TYPE DFC_rbr_outK62SCG : STRUCT
  DTC : UDINT := 16#043C00;
  DFCid : UINT := 682;
  debounceMethod : USINT := TIME_UP_DOWN;
END_STRUCT;
END_TYPE

TYPE DFC_rbr_outK62OR : STRUCT
  DTC : UDINT := 16#043A00;
  DFCid : UINT := 680;
  debounceMethod : USINT := TIME_UP_DOWN;
END_STRUCT;
END_TYPE

TYPE DFC_rbr_safoutChnl1 : STRUCT
  DTC : UDINT := 16#200800;
  DFCid : UINT := 1073;
  debounceMethod : USINT := NO_DEBOUNCE;
END_STRUCT;
END_TYPE

TYPE DFC_rbr_safoutChnl2 : STRUCT
  DTC : UDINT := 16#200900;
  DFCid : UINT := 1103;
  debounceMethod : USINT := NO_DEBOUNCE;
END_STRUCT;
END_TYPE

TYPE DFC_rbr_safoutChnl3 : STRUCT
  DTC : UDINT := 16#200A00;
  DFCid : UINT := 1106;
  debounceMethod : USINT := NO_DEBOUNCE;
END_STRUCT;
END_TYPE

TYPE DFC_rbr_safoutChnl4 : STRUCT
  DTC : UDINT := 16#200B00;
  DFCid : UINT := 1109;
  debounceMethod : USINT := NO_DEBOUNCE;
END_STRUCT;
END_TYPE

TYPE DFC_rbr_safoutChnl5 : STRUCT
  DTC : UDINT := 16#200C00;
  DFCid : UINT := 1112;
  debounceMethod : USINT := NO_DEBOUNCE;
END_STRUCT;
END_TYPE

TYPE DFC_rbr_safoutChnl6 : STRUCT
  DTC : UDINT := 16#201900;
  DFCid : UINT := 1115;
  debounceMethod : USINT := NO_DEBOUNCE;
END_STRUCT;
END_TYPE

TYPE DFC_rbr_safoutChnl7 : STRUCT
  DTC : UDINT := 16#201A00;
  DFCid : UINT := 1118;
  debounceMethod : USINT := NO_DEBOUNCE;
END_STRUCT;
END_TYPE

TYPE DFC_rbr_safoutChnl8 : STRUCT
  DTC : UDINT := 16#201B00;
  DFCid : UINT := 1121;
  debounceMethod : USINT := NO_DEBOUNCE;
END_STRUCT;
END_TYPE

TYPE DFC_rbr_safoutChnl9 : STRUCT
  DTC : UDINT := 16#201C00;
  DFCid : UINT := 1124;
  debounceMethod : USINT := NO_DEBOUNCE;
END_STRUCT;
END_TYPE

TYPE DFC_rbr_safoutChnl10 : STRUCT
  DTC : UDINT := 16#201D00;
  DFCid : UINT := 1074;
  debounceMethod : USINT := NO_DEBOUNCE;
END_STRUCT;
END_TYPE

TYPE DFC_rbr_safoutChnl11 : STRUCT
  DTC : UDINT := 16#201E00;
  DFCid : UINT := 1077;
  debounceMethod : USINT := NO_DEBOUNCE;
END_STRUCT;
END_TYPE

TYPE DFC_rbr_safoutChnl12 : STRUCT
  DTC : UDINT := 16#201F00;
  DFCid : UINT := 1080;
  debounceMethod : USINT := NO_DEBOUNCE;
END_STRUCT;
END_TYPE

TYPE DFC_rbr_safoutChnl13 : STRUCT
  DTC : UDINT := 16#202000;
  DFCid : UINT := 1083;
  debounceMethod : USINT := NO_DEBOUNCE;
END_STRUCT;
END_TYPE

TYPE DFC_rbr_safoutChnl14 : STRUCT
  DTC : UDINT := 16#202100;
  DFCid : UINT := 1086;
  debounceMethod : USINT := NO_DEBOUNCE;
END_STRUCT;
END_TYPE

TYPE DFC_rbr_safoutChnl15 : STRUCT
  DTC : UDINT := 16#202200;
  DFCid : UINT := 1089;
  debounceMethod : USINT := NO_DEBOUNCE;
END_STRUCT;
END_TYPE

TYPE DFC_rbr_safoutChnl16 : STRUCT
  DTC : UDINT := 16#202300;
  DFCid : UINT := 1092;
  debounceMethod : USINT := NO_DEBOUNCE;
END_STRUCT;
END_TYPE

TYPE DFC_rbr_safoutChnl17 : STRUCT
  DTC : UDINT := 16#202400;
  DFCid : UINT := 1095;
  debounceMethod : USINT := NO_DEBOUNCE;
END_STRUCT;
END_TYPE

TYPE DFC_rbr_safoutChnl18 : STRUCT
  DTC : UDINT := 16#202500;
  DFCid : UINT := 1098;
  debounceMethod : USINT := NO_DEBOUNCE;
END_STRUCT;
END_TYPE

TYPE DFC_rbr_safoutChnl6Dev : STRUCT
  DTC : UDINT := 16#202600;
  DFCid : UINT := 1116;
  debounceMethod : USINT := NO_DEBOUNCE;
END_STRUCT;
END_TYPE

TYPE DFC_rbr_safoutChnl7Dev : STRUCT
  DTC : UDINT := 16#202700;
  DFCid : UINT := 1119;
  debounceMethod : USINT := NO_DEBOUNCE;
END_STRUCT;
END_TYPE

TYPE DFC_rbr_safoutChnl8Dev : STRUCT
  DTC : UDINT := 16#202800;
  DFCid : UINT := 1122;
  debounceMethod : USINT := NO_DEBOUNCE;
END_STRUCT;
END_TYPE

TYPE DFC_rbr_safoutChnl9Dev : STRUCT
  DTC : UDINT := 16#202900;
  DFCid : UINT := 1125;
  debounceMethod : USINT := NO_DEBOUNCE;
END_STRUCT;
END_TYPE

TYPE DFC_rbr_safoutChnl10Dev : STRUCT
  DTC : UDINT := 16#202A00;
  DFCid : UINT := 1075;
  debounceMethod : USINT := NO_DEBOUNCE;
END_STRUCT;
END_TYPE

TYPE DFC_rbr_safoutChnl11Dev : STRUCT
  DTC : UDINT := 16#202B00;
  DFCid : UINT := 1078;
  debounceMethod : USINT := NO_DEBOUNCE;
END_STRUCT;
END_TYPE

TYPE DFC_rbr_safoutChnl12Dev : STRUCT
  DTC : UDINT := 16#202C00;
  DFCid : UINT := 1081;
  debounceMethod : USINT := NO_DEBOUNCE;
END_STRUCT;
END_TYPE

TYPE DFC_rbr_safoutChnl13Dev : STRUCT
  DTC : UDINT := 16#202D00;
  DFCid : UINT := 1084;
  debounceMethod : USINT := NO_DEBOUNCE;
END_STRUCT;
END_TYPE

TYPE DFC_rbr_safoutChnl14Dev : STRUCT
  DTC : UDINT := 16#202E00;
  DFCid : UINT := 1087;
  debounceMethod : USINT := NO_DEBOUNCE;
END_STRUCT;
END_TYPE

TYPE DFC_rbr_safoutChnl15Dev : STRUCT
  DTC : UDINT := 16#202F00;
  DFCid : UINT := 1090;
  debounceMethod : USINT := NO_DEBOUNCE;
END_STRUCT;
END_TYPE

TYPE DFC_rbr_safoutChnl16Dev : STRUCT
  DTC : UDINT := 16#203000;
  DFCid : UINT := 1093;
  debounceMethod : USINT := NO_DEBOUNCE;
END_STRUCT;
END_TYPE

TYPE DFC_rbr_safoutChnl17Dev : STRUCT
  DTC : UDINT := 16#203100;
  DFCid : UINT := 1096;
  debounceMethod : USINT := NO_DEBOUNCE;
END_STRUCT;
END_TYPE

TYPE DFC_rbr_safoutChnl18Dev : STRUCT
  DTC : UDINT := 16#203200;
  DFCid : UINT := 1099;
  debounceMethod : USINT := NO_DEBOUNCE;
END_STRUCT;
END_TYPE

TYPE DFC_rbr_safoutChnl1OR : STRUCT
  DTC : UDINT := 16#200D00;
  DFCid : UINT := 1102;
  debounceMethod : USINT := NO_DEBOUNCE;
END_STRUCT;
END_TYPE

TYPE DFC_rbr_safoutChnl2OR : STRUCT
  DTC : UDINT := 16#200E00;
  DFCid : UINT := 1105;
  debounceMethod : USINT := NO_DEBOUNCE;
END_STRUCT;
END_TYPE

TYPE DFC_rbr_safoutChnl3OR : STRUCT
  DTC : UDINT := 16#200F00;
  DFCid : UINT := 1108;
  debounceMethod : USINT := NO_DEBOUNCE;
END_STRUCT;
END_TYPE

TYPE DFC_rbr_safoutChnl4OR : STRUCT
  DTC : UDINT := 16#201100;
  DFCid : UINT := 1111;
  debounceMethod : USINT := NO_DEBOUNCE;
END_STRUCT;
END_TYPE

TYPE DFC_rbr_safoutChnl5OR : STRUCT
  DTC : UDINT := 16#201200;
  DFCid : UINT := 1114;
  debounceMethod : USINT := NO_DEBOUNCE;
END_STRUCT;
END_TYPE

TYPE DFC_rbr_safoutChnl6OR : STRUCT
  DTC : UDINT := 16#203300;
  DFCid : UINT := 1117;
  debounceMethod : USINT := NO_DEBOUNCE;
END_STRUCT;
END_TYPE

TYPE DFC_rbr_safoutChnl7OR : STRUCT
  DTC : UDINT := 16#203400;
  DFCid : UINT := 1120;
  debounceMethod : USINT := NO_DEBOUNCE;
END_STRUCT;
END_TYPE

TYPE DFC_rbr_safoutChnl8OR : STRUCT
  DTC : UDINT := 16#203500;
  DFCid : UINT := 1123;
  debounceMethod : USINT := NO_DEBOUNCE;
END_STRUCT;
END_TYPE

TYPE DFC_rbr_safoutChnl9OR : STRUCT
  DTC : UDINT := 16#203600;
  DFCid : UINT := 1126;
  debounceMethod : USINT := NO_DEBOUNCE;
END_STRUCT;
END_TYPE

TYPE DFC_rbr_safoutChnl10OR : STRUCT
  DTC : UDINT := 16#203700;
  DFCid : UINT := 1076;
  debounceMethod : USINT := NO_DEBOUNCE;
END_STRUCT;
END_TYPE

TYPE DFC_rbr_safoutChnl11OR : STRUCT
  DTC : UDINT := 16#203800;
  DFCid : UINT := 1079;
  debounceMethod : USINT := NO_DEBOUNCE;
END_STRUCT;
END_TYPE

TYPE DFC_rbr_safoutChnl12OR : STRUCT
  DTC : UDINT := 16#203900;
  DFCid : UINT := 1082;
  debounceMethod : USINT := NO_DEBOUNCE;
END_STRUCT;
END_TYPE

TYPE DFC_rbr_safoutChnl13OR : STRUCT
  DTC : UDINT := 16#203A00;
  DFCid : UINT := 1085;
  debounceMethod : USINT := NO_DEBOUNCE;
END_STRUCT;
END_TYPE

TYPE DFC_rbr_safoutChnl14OR : STRUCT
  DTC : UDINT := 16#203B00;
  DFCid : UINT := 1088;
  debounceMethod : USINT := NO_DEBOUNCE;
END_STRUCT;
END_TYPE

TYPE DFC_rbr_safoutChnl15OR : STRUCT
  DTC : UDINT := 16#203C00;
  DFCid : UINT := 1091;
  debounceMethod : USINT := NO_DEBOUNCE;
END_STRUCT;
END_TYPE

TYPE DFC_rbr_safoutChnl16OR : STRUCT
  DTC : UDINT := 16#203D00;
  DFCid : UINT := 1094;
  debounceMethod : USINT := NO_DEBOUNCE;
END_STRUCT;
END_TYPE

TYPE DFC_rbr_safoutChnl17OR : STRUCT
  DTC : UDINT := 16#203E00;
  DFCid : UINT := 1097;
  debounceMethod : USINT := NO_DEBOUNCE;
END_STRUCT;
END_TYPE

TYPE DFC_rbr_safoutChnl18OR : STRUCT
  DTC : UDINT := 16#203F00;
  DFCid : UINT := 1100;
  debounceMethod : USINT := NO_DEBOUNCE;
END_STRUCT;
END_TYPE

TYPE DFC_rbr_safoutCfg : STRUCT
  DTC : UDINT := 16#200100;
  DFCid : UINT := 1072;
  debounceMethod : USINT := NO_DEBOUNCE;
END_STRUCT;
END_TYPE

TYPE DFC_rbr_safout : STRUCT
  DTC : UDINT := 16#200200;
  DFCid : UINT := 1071;
  debounceMethod : USINT := NO_DEBOUNCE;
END_STRUCT;
END_TYPE

TYPE DFC_rbr_safoutGetStatus : STRUCT
  DTC : UDINT := 16#200300;
  DFCid : UINT := 1128;
  debounceMethod : USINT := NO_DEBOUNCE;
END_STRUCT;
END_TYPE

TYPE DFC_rbr_safoutDevError : STRUCT
  DTC : UDINT := 16#201800;
  DFCid : UINT := 1127;
  debounceMethod : USINT := NO_DEBOUNCE;
END_STRUCT;
END_TYPE

TYPE DFC_rbr_safoutResetError : STRUCT
  DTC : UDINT := 16#200400;
  DFCid : UINT := 1130;
  debounceMethod : USINT := NO_DEBOUNCE;
END_STRUCT;
END_TYPE

TYPE DFC_rbr_safoutIgnoreError : STRUCT
  DTC : UDINT := 16#200500;
  DFCid : UINT := 1129;
  debounceMethod : USINT := NO_DEBOUNCE;
END_STRUCT;
END_TYPE

TYPE DFC_rbr_safoutUnlock : STRUCT
  DTC : UDINT := 16#200600;
  DFCid : UINT := 1131;
  debounceMethod : USINT := NO_DEBOUNCE;
END_STRUCT;
END_TYPE

TYPE DFC_rbr_outDo : STRUCT
  DTC : UDINT := 16#048300;
  DFCid : UINT := 1025;
  debounceMethod : USINT := NO_DEBOUNCE;
END_STRUCT;
END_TYPE

TYPE DFC_rbr_outDoGetCurrent : STRUCT
  DTC : UDINT := 16#048400;
  DFCid : UINT := 1028;
  debounceMethod : USINT := NO_DEBOUNCE;
END_STRUCT;
END_TYPE

TYPE DFC_rbr_outPod : STRUCT
  DTC : UDINT := 16#048B00;
  DFCid : UINT := 1067;
  debounceMethod : USINT := NO_DEBOUNCE;
END_STRUCT;
END_TYPE

TYPE DFC_rbr_outPodCfg : STRUCT
  DTC : UDINT := 16#048C00;
  DFCid : UINT := 1068;
  debounceMethod : USINT := NO_DEBOUNCE;
END_STRUCT;
END_TYPE

TYPE DFC_rbr_outPodCfgPeriod : STRUCT
  DTC : UDINT := 16#048D00;
  DFCid : UINT := 1069;
  debounceMethod : USINT := NO_DEBOUNCE;
END_STRUCT;
END_TYPE

TYPE DFC_rbr_outPoc : STRUCT
  DTC : UDINT := 16#048600;
  DFCid : UINT := 1063;
  debounceMethod : USINT := NO_DEBOUNCE;
END_STRUCT;
END_TYPE

TYPE DFC_rbr_outPocCfg : STRUCT
  DTC : UDINT := 16#048800;
  DFCid : UINT := 1064;
  debounceMethod : USINT := NO_DEBOUNCE;
END_STRUCT;
END_TYPE

TYPE DFC_rbr_outPoCfg : STRUCT
  DTC : UDINT := 16#048700;
  DFCid : UINT := 1056;
  debounceMethod : USINT := NO_DEBOUNCE;
END_STRUCT;
END_TYPE

TYPE DFC_rbr_outPocCfgPI : STRUCT
  DTC : UDINT := 16#048A00;
  DFCid : UINT := 1066;
  debounceMethod : USINT := NO_DEBOUNCE;
END_STRUCT;
END_TYPE

TYPE DFC_rbr_outPocCfgDither : STRUCT
  DTC : UDINT := 16#048900;
  DFCid : UINT := 1065;
  debounceMethod : USINT := NO_DEBOUNCE;
END_STRUCT;
END_TYPE

TYPE DFC_rbr_outPoGetCurrent : STRUCT
  DTC : UDINT := 16#048E00;
  DFCid : UINT := 1060;
  debounceMethod : USINT := NO_DEBOUNCE;
END_STRUCT;
END_TYPE

TYPE DFC_rbr_outAov : STRUCT
  DTC : UDINT := 16#048000;
  DFCid : UINT := 1019;
  debounceMethod : USINT := NO_DEBOUNCE;
END_STRUCT;
END_TYPE

TYPE DFC_rbr_outAovCfg : STRUCT
  DTC : UDINT := 16#048100;
  DFCid : UINT := 1020;
  debounceMethod : USINT := NO_DEBOUNCE;
END_STRUCT;
END_TYPE

TYPE DFC_rbr_outAovCfgPI : STRUCT
  DTC : UDINT := 16#14D700;
  DFCid : UINT := 1021;
  debounceMethod : USINT := NO_DEBOUNCE;
END_STRUCT;
END_TYPE

TYPE DFC_rbr_outAovGetVoltage : STRUCT
  DTC : UDINT := 16#048200;
  DFCid : UINT := 1023;
  debounceMethod : USINT := NO_DEBOUNCE;
END_STRUCT;
END_TYPE

TYPE DFC_rbr_outDoGetStatus : STRUCT
  DTC : UDINT := 16#048F00;
  DFCid : UINT := 1029;
  debounceMethod : USINT := NO_DEBOUNCE;
END_STRUCT;
END_TYPE

TYPE DFC_rbr_outDoResetError : STRUCT
  DTC : UDINT := 16#049000;
  DFCid : UINT := 1030;
  debounceMethod : USINT := NO_DEBOUNCE;
END_STRUCT;
END_TYPE

TYPE DFC_rbr_outPo : STRUCT
  DTC : UDINT := 16#049100;
  DFCid : UINT := 1055;
  debounceMethod : USINT := NO_DEBOUNCE;
END_STRUCT;
END_TYPE

TYPE DFC_rbr_outPoCfgPeriod : STRUCT
  DTC : UDINT := 16#049200;
  DFCid : UINT := 1057;
  debounceMethod : USINT := NO_DEBOUNCE;
END_STRUCT;
END_TYPE

TYPE DFC_rbr_outPoGetStatus : STRUCT
  DTC : UDINT := 16#049300;
  DFCid : UINT := 1061;
  debounceMethod : USINT := NO_DEBOUNCE;
END_STRUCT;
END_TYPE

TYPE DFC_rbr_outPoResetError : STRUCT
  DTC : UDINT := 16#049400;
  DFCid : UINT := 1062;
  debounceMethod : USINT := NO_DEBOUNCE;
END_STRUCT;
END_TYPE

TYPE DFC_rbr_outAovGetStatus : STRUCT
  DTC : UDINT := 16#049500;
  DFCid : UINT := 1022;
  debounceMethod : USINT := NO_DEBOUNCE;
END_STRUCT;
END_TYPE

TYPE DFC_rbr_outAovResetError : STRUCT
  DTC : UDINT := 16#049600;
  DFCid : UINT := 1024;
  debounceMethod : USINT := NO_DEBOUNCE;
END_STRUCT;
END_TYPE

TYPE DFC_rbr_sysAiv : STRUCT
  DTC : UDINT := 16#010100;
  DFCid : UINT := 1146;
  debounceMethod : USINT := NO_DEBOUNCE;
END_STRUCT;
END_TYPE

TYPE DFC_rbr_memFlsCfgShr : STRUCT
  DTC : UDINT := 16#060900;
  DFCid : UINT := 953;
  debounceMethod : USINT := NO_DEBOUNCE;
END_STRUCT;
END_TYPE

TYPE DFC_rbr_sysDo : STRUCT
  DTC : UDINT := 16#010200;
  DFCid : UINT := 1148;
  debounceMethod : USINT := NO_DEBOUNCE;
END_STRUCT;
END_TYPE

TYPE DFC_rbr_sysGetVss : STRUCT
  DTC : UDINT := 16#010600;
  DFCid : UINT := 1149;
  debounceMethod : USINT := NO_DEBOUNCE;
END_STRUCT;
END_TYPE

TYPE DFC_rbr_sysDi : STRUCT
  DTC : UDINT := 16#010300;
  DFCid : UINT := 1147;
  debounceMethod : USINT := NO_DEBOUNCE;
END_STRUCT;
END_TYPE

TYPE DFC_rbr_sysAit : STRUCT
  DTC : UDINT := 16#010400;
  DFCid : UINT := 1145;
  debounceMethod : USINT := NO_DEBOUNCE;
END_STRUCT;
END_TYPE

TYPE DFC_rbr_sysSetVss : STRUCT
  DTC : UDINT := 16#010500;
  DFCid : UINT := 1153;
  debounceMethod : USINT := NO_DEBOUNCE;
END_STRUCT;
END_TYPE

TYPE DFC_rbr_outPoDisable : STRUCT
  DTC : UDINT := 16#049800;
  DFCid : UINT := 1059;
  debounceMethod : USINT := NO_DEBOUNCE;
END_STRUCT;
END_TYPE

TYPE DFC_rbr_safout_cfgDiag : STRUCT
  DTC : UDINT := 16#200700;
  DFCid : UINT := 1132;
  debounceMethod : USINT := NO_DEBOUNCE;
END_STRUCT;
END_TYPE

TYPE DFC_rbr_outDoDisable : STRUCT
  DTC : UDINT := 16#049700;
  DFCid : UINT := 1027;
  debounceMethod : USINT := NO_DEBOUNCE;
END_STRUCT;
END_TYPE

TYPE DFC_rbr_sysOperHrIntegrityErr : STRUCT
  DTC : UDINT := 16#010A00;
  DFCid : UINT := 1151;
  debounceMethod : USINT := NO_DEBOUNCE;
END_STRUCT;
END_TYPE

TYPE DFC_rbr_sysOperHrsSaturated : STRUCT
  DTC : UDINT := 16#010B00;
  DFCid : UINT := 1152;
  debounceMethod : USINT := NO_DEBOUNCE;
END_STRUCT;
END_TYPE

TYPE DFC_rbr_mo_INHLatch : STRUCT
  DTC : UDINT := 16#082200;
  DFCid : UINT := 968;
  debounceMethod : USINT := NO_DEBOUNCE;
END_STRUCT;
END_TYPE

TYPE DFC_rbr_mo_INH : STRUCT
  DTC : UDINT := 16#082100;
  DFCid : UINT := 967;
  debounceMethod : USINT := NO_DEBOUNCE;
END_STRUCT;
END_TYPE

TYPE DFC_rbr_memReadSystemError : STRUCT
  DTC : UDINT := 16#060800;
  DFCid : UINT := 961;
  debounceMethod : USINT := NO_DEBOUNCE;
END_STRUCT;
END_TYPE

TYPE DFC_rbr_memReadCalibInputError : STRUCT
  DTC : UDINT := 16#060A00;
  DFCid : UINT := 959;
  debounceMethod : USINT := NO_DEBOUNCE;
END_STRUCT;
END_TYPE

TYPE DFC_rbr_memReadCalibOuputError : STRUCT
  DTC : UDINT := 16#060B00;
  DFCid : UINT := 960;
  debounceMethod : USINT := NO_DEBOUNCE;
END_STRUCT;
END_TYPE

TYPE DFC_rbr_memReadApi2Error : STRUCT
  DTC : UDINT := 16#060600;
  DFCid : UINT := 957;
  debounceMethod : USINT := NO_DEBOUNCE;
END_STRUCT;
END_TYPE

TYPE DFC_rbr_memReadApi1Error : STRUCT
  DTC : UDINT := 16#060500;
  DFCid : UINT := 956;
  debounceMethod : USINT := NO_DEBOUNCE;
END_STRUCT;
END_TYPE

TYPE DFC_rbr_memMarkBlock : STRUCT
  DTC : UDINT := 16#060400;
  DFCid : UINT := 955;
  debounceMethod : USINT := NO_DEBOUNCE;
END_STRUCT;
END_TYPE

TYPE DFC_rbr_safoutChnl3Dev : STRUCT
  DTC : UDINT := 16#201500;
  DFCid : UINT := 1107;
  debounceMethod : USINT := NO_DEBOUNCE;
END_STRUCT;
END_TYPE

TYPE DFC_rbr_safoutChnl5Dev : STRUCT
  DTC : UDINT := 16#201700;
  DFCid : UINT := 1113;
  debounceMethod : USINT := NO_DEBOUNCE;
END_STRUCT;
END_TYPE

TYPE DFC_rbr_safoutChnl4Dev : STRUCT
  DTC : UDINT := 16#201600;
  DFCid : UINT := 1110;
  debounceMethod : USINT := NO_DEBOUNCE;
END_STRUCT;
END_TYPE

TYPE DFC_rbr_safoutChnl2Dev : STRUCT
  DTC : UDINT := 16#201400;
  DFCid : UINT := 1104;
  debounceMethod : USINT := NO_DEBOUNCE;
END_STRUCT;
END_TYPE

TYPE DFC_rbr_safoutChnl1Dev : STRUCT
  DTC : UDINT := 16#201300;
  DFCid : UINT := 1101;
  debounceMethod : USINT := NO_DEBOUNCE;
END_STRUCT;
END_TYPE

TYPE DFC_rbr_outPoCfgPwrLs : STRUCT
  DTC : UDINT := 16#049900;
  DFCid : UINT := 1058;
  debounceMethod : USINT := NO_DEBOUNCE;
END_STRUCT;
END_TYPE

TYPE DFC_rbr_lin_wakeUp : STRUCT
  DTC : UDINT := 16#210000;
  DFCid : UINT := 952;
  debounceMethod : USINT := NO_DEBOUNCE;
END_STRUCT;
END_TYPE

TYPE DFC_rbr_lin_gotoSleep : STRUCT
  DTC : UDINT := 16#210200;
  DFCid : UINT := 950;
  debounceMethod : USINT := NO_DEBOUNCE;
END_STRUCT;
END_TYPE

TYPE DFC_rbr_lin_getStatus : STRUCT
  DTC : UDINT := 16#210300;
  DFCid : UINT := 949;
  debounceMethod : USINT := NO_DEBOUNCE;
END_STRUCT;
END_TYPE

TYPE DFC_rbr_lin_scheduleRequest : STRUCT
  DTC : UDINT := 16#210100;
  DFCid : UINT := 951;
  debounceMethod : USINT := NO_DEBOUNCE;
END_STRUCT;
END_TYPE

TYPE DFC_rbr_lin_SendSignal : STRUCT
  DTC : UDINT := 16#210400;
  DFCid : UINT := 948;
  debounceMethod : USINT := NO_DEBOUNCE;
END_STRUCT;
END_TYPE

TYPE DFC_rbr_inPhaseGetStatus : STRUCT
  DTC : UDINT := 16#039F00;
  DFCid : UINT := 897;
  debounceMethod : USINT := NO_DEBOUNCE;
END_STRUCT;
END_TYPE

TYPE DFC_rbr_inPhaseResetCounter : STRUCT
  DTC : UDINT := 16#03A000;
  DFCid : UINT := 898;
  debounceMethod : USINT := NO_DEBOUNCE;
END_STRUCT;
END_TYPE

TYPE DFC_rbr_inPhase : STRUCT
  DTC : UDINT := 16#039E00;
  DFCid : UINT := 896;
  debounceMethod : USINT := NO_DEBOUNCE;
END_STRUCT;
END_TYPE

TYPE DFC_rbr_inFi_Buffered : STRUCT
  DTC : UDINT := 16#135200;
  DFCid : UINT := 895;
  debounceMethod : USINT := NO_DEBOUNCE;
END_STRUCT;
END_TYPE

TYPE DFC_rbr_secGetLevel : STRUCT
  DTC : UDINT := 16#220200;
  DFCid : UINT := 1137;
  debounceMethod : USINT := NO_DEBOUNCE;
END_STRUCT;
END_TYPE

TYPE DFC_rbr_secSetLevel : STRUCT
  DTC : UDINT := 16#220300;
  DFCid : UINT := 1144;
  debounceMethod : USINT := NO_DEBOUNCE;
END_STRUCT;
END_TYPE

TYPE DFC_rbr_secSaveSecret : STRUCT
  DTC : UDINT := 16#220100;
  DFCid : UINT := 1143;
  debounceMethod : USINT := NO_DEBOUNCE;
END_STRUCT;
END_TYPE

TYPE DFC_rbr_secGetSeed : STRUCT
  DTC : UDINT := 16#220000;
  DFCid : UINT := 1139;
  debounceMethod : USINT := NO_DEBOUNCE;
END_STRUCT;
END_TYPE

TYPE DFC_rbr_secIsRequestAllowed : STRUCT
  DTC : UDINT := 16#220700;
  DFCid : UINT := 1141;
  debounceMethod : USINT := NO_DEBOUNCE;
END_STRUCT;
END_TYPE

TYPE DFC_rbr_secGetRnd : STRUCT
  DTC : UDINT := 16#220600;
  DFCid : UINT := 1138;
  debounceMethod : USINT := NO_DEBOUNCE;
END_STRUCT;
END_TYPE

TYPE DFC_rbr_secEvalRespKey : STRUCT
  DTC : UDINT := 16#220500;
  DFCid : UINT := 1135;
  debounceMethod : USINT := NO_DEBOUNCE;
END_STRUCT;
END_TYPE

TYPE DFC_rbr_secResetLevel : STRUCT
  DTC : UDINT := 16#220400;
  DFCid : UINT := 1142;
  debounceMethod : USINT := NO_DEBOUNCE;
END_STRUCT;
END_TYPE

TYPE DFC_rbr_lin_ReceiveSignal : STRUCT
  DTC : UDINT := 16#210500;
  DFCid : UINT := 947;
  debounceMethod : USINT := NO_DEBOUNCE;
END_STRUCT;
END_TYPE

TYPE DFC_rbr_sys_coreload : STRUCT
  DTC : UDINT := 16#010900;
  DFCid : UINT := 1154;
  debounceMethod : USINT := NO_DEBOUNCE;
END_STRUCT;
END_TYPE

TYPE DFC_rbr_sys_taskload : STRUCT
  DTC : UDINT := 16#010800;
  DFCid : UINT := 1155;
  debounceMethod : USINT := NO_DEBOUNCE;
END_STRUCT;
END_TYPE

TYPE DFC_rbr_dsmDTCJ1939 : STRUCT
  DTC : UDINT := 16#071000;
  DFCid : UINT := 868;
  debounceMethod : USINT := NO_DEBOUNCE;
END_STRUCT;
END_TYPE

TYPE DFC_rbr_sysInit : STRUCT
  DTC : UDINT := 16#010700;
  DFCid : UINT := 1150;
  debounceMethod : USINT := NO_DEBOUNCE;
END_STRUCT;
END_TYPE

TYPE DFC_rbr_outK07Unintended : STRUCT
  DTC : UDINT := 16#14CB00;
  DFCid : UINT := 1032;
  debounceMethod : USINT := NO_DEBOUNCE;
END_STRUCT;
END_TYPE

TYPE DFC_rbr_outK09Unintended : STRUCT
  DTC : UDINT := 16#14CD00;
  DFCid : UINT := 1036;
  debounceMethod : USINT := NO_DEBOUNCE;
END_STRUCT;
END_TYPE

TYPE DFC_rbr_outK73Unintended : STRUCT
  DTC : UDINT := 16#14D600;
  DFCid : UINT := 1054;
  debounceMethod : USINT := NO_DEBOUNCE;
END_STRUCT;
END_TYPE

TYPE DFC_rbr_outK08Unintended : STRUCT
  DTC : UDINT := 16#14CC00;
  DFCid : UINT := 1034;
  debounceMethod : USINT := NO_DEBOUNCE;
END_STRUCT;
END_TYPE

TYPE DFC_rbr_outK29Unintended : STRUCT
  DTC : UDINT := 16#14D400;
  DFCid : UINT := 1050;
  debounceMethod : USINT := NO_DEBOUNCE;
END_STRUCT;
END_TYPE

TYPE DFC_rbr_outK17Unintended : STRUCT
  DTC : UDINT := 16#14D300;
  DFCid : UINT := 1048;
  debounceMethod : USINT := NO_DEBOUNCE;
END_STRUCT;
END_TYPE

TYPE DFC_rbr_outK16Unintended : STRUCT
  DTC : UDINT := 16#14D200;
  DFCid : UINT := 1046;
  debounceMethod : USINT := NO_DEBOUNCE;
END_STRUCT;
END_TYPE

TYPE DFC_rbr_outK14Unintended : STRUCT
  DTC : UDINT := 16#14D000;
  DFCid : UINT := 1042;
  debounceMethod : USINT := NO_DEBOUNCE;
END_STRUCT;
END_TYPE

TYPE DFC_rbr_outK15Unintended : STRUCT
  DTC : UDINT := 16#14D100;
  DFCid : UINT := 1044;
  debounceMethod : USINT := NO_DEBOUNCE;
END_STRUCT;
END_TYPE

TYPE DFC_rbr_outK51Unintended : STRUCT
  DTC : UDINT := 16#14D500;
  DFCid : UINT := 1052;
  debounceMethod : USINT := NO_DEBOUNCE;
END_STRUCT;
END_TYPE

TYPE DFC_rbr_outK12Unintended : STRUCT
  DTC : UDINT := 16#14CE00;
  DFCid : UINT := 1038;
  debounceMethod : USINT := NO_DEBOUNCE;
END_STRUCT;
END_TYPE

TYPE DFC_rbr_outK13Unintended : STRUCT
  DTC : UDINT := 16#14CF00;
  DFCid : UINT := 1040;
  debounceMethod : USINT := NO_DEBOUNCE;
END_STRUCT;
END_TYPE

TYPE DFC_rbr_outA32Unintended : STRUCT
  DTC : UDINT := 16#14C000;
  DFCid : UINT := 998;
  debounceMethod : USINT := NO_DEBOUNCE;
END_STRUCT;
END_TYPE

TYPE DFC_rbr_outA47Unintended : STRUCT
  DTC : UDINT := 16#14C500;
  DFCid : UINT := 1008;
  debounceMethod : USINT := NO_DEBOUNCE;
END_STRUCT;
END_TYPE

TYPE DFC_rbr_outA31Unintended : STRUCT
  DTC : UDINT := 16#14BF00;
  DFCid : UINT := 996;
  debounceMethod : USINT := NO_DEBOUNCE;
END_STRUCT;
END_TYPE

TYPE DFC_rbr_outA48Unintended : STRUCT
  DTC : UDINT := 16#14C600;
  DFCid : UINT := 1010;
  debounceMethod : USINT := NO_DEBOUNCE;
END_STRUCT;
END_TYPE

TYPE DFC_rbr_outA46Unintended : STRUCT
  DTC : UDINT := 16#14C400;
  DFCid : UINT := 1006;
  debounceMethod : USINT := NO_DEBOUNCE;
END_STRUCT;
END_TYPE

TYPE DFC_rbr_outA33Unintended : STRUCT
  DTC : UDINT := 16#14C100;
  DFCid : UINT := 1000;
  debounceMethod : USINT := NO_DEBOUNCE;
END_STRUCT;
END_TYPE

TYPE DFC_rbr_outA19Unintended : STRUCT
  DTC : UDINT := 16#14BD00;
  DFCid : UINT := 992;
  debounceMethod : USINT := NO_DEBOUNCE;
END_STRUCT;
END_TYPE

TYPE DFC_rbr_outA05Unintended : STRUCT
  DTC : UDINT := 16#14B600;
  DFCid : UINT := 978;
  debounceMethod : USINT := NO_DEBOUNCE;
END_STRUCT;
END_TYPE

TYPE DFC_rbr_outA20Unintended : STRUCT
  DTC : UDINT := 16#14BE00;
  DFCid : UINT := 994;
  debounceMethod : USINT := NO_DEBOUNCE;
END_STRUCT;
END_TYPE

TYPE DFC_rbr_outA03Unintended : STRUCT
  DTC : UDINT := 16#14B400;
  DFCid : UINT := 974;
  debounceMethod : USINT := NO_DEBOUNCE;
END_STRUCT;
END_TYPE

TYPE DFC_rbr_outA18Unintended : STRUCT
  DTC : UDINT := 16#14BC00;
  DFCid : UINT := 990;
  debounceMethod : USINT := NO_DEBOUNCE;
END_STRUCT;
END_TYPE

TYPE DFC_rbr_outA04Unintended : STRUCT
  DTC : UDINT := 16#14B500;
  DFCid : UINT := 976;
  debounceMethod : USINT := NO_DEBOUNCE;
END_STRUCT;
END_TYPE

TYPE DFC_rbr_outA34Unintended : STRUCT
  DTC : UDINT := 16#14C200;
  DFCid : UINT := 1002;
  debounceMethod : USINT := NO_DEBOUNCE;
END_STRUCT;
END_TYPE

TYPE DFC_rbr_outA51Unintended : STRUCT
  DTC : UDINT := 16#14C700;
  DFCid : UINT := 1012;
  debounceMethod : USINT := NO_DEBOUNCE;
END_STRUCT;
END_TYPE

TYPE DFC_rbr_outA35Unintended : STRUCT
  DTC : UDINT := 16#14C300;
  DFCid : UINT := 1004;
  debounceMethod : USINT := NO_DEBOUNCE;
END_STRUCT;
END_TYPE

TYPE DFC_rbr_outA53Unintended : STRUCT
  DTC : UDINT := 16#14C900;
  DFCid : UINT := 1016;
  debounceMethod : USINT := NO_DEBOUNCE;
END_STRUCT;
END_TYPE

TYPE DFC_rbr_outA52Unintended : STRUCT
  DTC : UDINT := 16#14C800;
  DFCid : UINT := 1014;
  debounceMethod : USINT := NO_DEBOUNCE;
END_STRUCT;
END_TYPE

TYPE DFC_rbr_outA54Unintended : STRUCT
  DTC : UDINT := 16#14CA00;
  DFCid : UINT := 1018;
  debounceMethod : USINT := NO_DEBOUNCE;
END_STRUCT;
END_TYPE

TYPE DFC_rbr_outA09Unintended : STRUCT
  DTC : UDINT := 16#14B900;
  DFCid : UINT := 984;
  debounceMethod : USINT := NO_DEBOUNCE;
END_STRUCT;
END_TYPE

TYPE DFC_rbr_outA02Unintended : STRUCT
  DTC : UDINT := 16#14B300;
  DFCid : UINT := 972;
  debounceMethod : USINT := NO_DEBOUNCE;
END_STRUCT;
END_TYPE

TYPE DFC_rbr_outA17Unintended : STRUCT
  DTC : UDINT := 16#14BB00;
  DFCid : UINT := 988;
  debounceMethod : USINT := NO_DEBOUNCE;
END_STRUCT;
END_TYPE

TYPE DFC_rbr_outA08Unintended : STRUCT
  DTC : UDINT := 16#14B800;
  DFCid : UINT := 982;
  debounceMethod : USINT := NO_DEBOUNCE;
END_STRUCT;
END_TYPE

TYPE DFC_rbr_outA07Unintended : STRUCT
  DTC : UDINT := 16#14B700;
  DFCid : UINT := 980;
  debounceMethod : USINT := NO_DEBOUNCE;
END_STRUCT;
END_TYPE

TYPE DFC_rbr_outA10Unintended : STRUCT
  DTC : UDINT := 16#14BA00;
  DFCid : UINT := 986;
  debounceMethod : USINT := NO_DEBOUNCE;
END_STRUCT;
END_TYPE

TYPE DFC_rbr_outDoCfgPwrLs : STRUCT
  DTC : UDINT := 16#14D800;
  DFCid : UINT := 1026;
  debounceMethod : USINT := NO_DEBOUNCE;
END_STRUCT;
END_TYPE

TYPE DFC_rbr_mo_memoryProtection_err : STRUCT
  DTC : UDINT := 16#083300;
  DFCid : UINT := 970;
  debounceMethod : USINT := NO_DEBOUNCE;
END_STRUCT;
END_TYPE

TYPE DFC_rbr_rsmFfiApiCallErr : STRUCT
  DTC : UDINT := 16#010C00;
  DFCid : UINT := 1070;
  debounceMethod : USINT := NO_DEBOUNCE;
END_STRUCT;
END_TYPE

TYPE DFC_rbr_isobusSftyCanTxErr : STRUCT
  DTC : UDINT := 16#051F00;
  DFCid : UINT := 946;
  debounceMethod : USINT := NO_DEBOUNCE;
END_STRUCT;
END_TYPE

TYPE DFC_rbr_dsmInitQueueOverflow : STRUCT
  DTC : UDINT := 16#071400;
  DFCid : UINT := 875;
  debounceMethod : USINT := NO_DEBOUNCE;
END_STRUCT;
END_TYPE

TYPE DFC_rbr_secAccessDenied_RC : STRUCT
  DTC : UDINT := 16#220B00;
  DFCid : UINT := 1133;
  debounceMethod : USINT := NO_DEBOUNCE;
END_STRUCT;
END_TYPE

TYPE DFC_rbr_secAccessDenied_WDBI : STRUCT
  DTC : UDINT := 16#220A00;
  DFCid : UINT := 1134;
  debounceMethod : USINT := NO_DEBOUNCE;
END_STRUCT;
END_TYPE

TYPE DFC_rbr_secFlashingFailure : STRUCT
  DTC : UDINT := 16#220900;
  DFCid : UINT := 1136;
  debounceMethod : USINT := NO_DEBOUNCE;
END_STRUCT;
END_TYPE

TYPE DFC_rbr_secInvalidPassword : STRUCT
  DTC : UDINT := 16#220800;
  DFCid : UINT := 1140;
  debounceMethod : USINT := NO_DEBOUNCE;
END_STRUCT;
END_TYPE

TYPE DFC_ComCntESP_05 : STRUCT
  DTC : UDINT := 16#102200;
END_STRUCT;
END_TYPE

TYPE DFC_MOXEMM_SMU_ALM3_1 : STRUCT
  DTC : UDINT := 16#108800;
  DFCid : UINT := 1237;
  debounceMethod : USINT := NATIVE;
END_STRUCT;
END_TYPE

TYPE DFC_MOXEMM_SMU_ALM3_2 : STRUCT
  DTC : UDINT := 16#108900;
  DFCid : UINT := 1242;
  debounceMethod : USINT := NATIVE;
END_STRUCT;
END_TYPE

TYPE DFC_ComCntESP_07 : STRUCT
  DTC : UDINT := 16#102300;
END_STRUCT;
END_TYPE

TYPE DFC_MOXEMM_SMU_ALM3_4 : STRUCT
  DTC : UDINT := 16#108A00;
  DFCid : UINT := 1245;
  debounceMethod : USINT := NATIVE;
END_STRUCT;
END_TYPE

TYPE DFC_MOXEMM_SMU_ALM3_5 : STRUCT
  DTC : UDINT := 16#108B00;
  DFCid : UINT := 1246;
  debounceMethod : USINT := NATIVE;
END_STRUCT;
END_TYPE

TYPE DFC_MOXEMM_SMU_ALM3_7 : STRUCT
  DTC : UDINT := 16#108C00;
  DFCid : UINT := 1247;
  debounceMethod : USINT := NATIVE;
END_STRUCT;
END_TYPE

TYPE DFC_MoXEMMHwLTRegMonTest : STRUCT
  DTC : UDINT := 16#10D400;
  DFCid : UINT := 1301;
  debounceMethod : USINT := NATIVE;
END_STRUCT;
END_TYPE

TYPE DFC_ComCntESP_02 : STRUCT
  DTC : UDINT := 16#102100;
END_STRUCT;
END_TYPE

TYPE DFC_DSMDummy : STRUCT
  DTC : UDINT := 16#100F00;
  DFCid : UINT := 720;
  debounceMethod : USINT := NO_DEBOUNCE;
END_STRUCT;
END_TYPE

TYPE DFC_MOXEMM_SMU_ALM2_22 : STRUCT
  DTC : UDINT := 16#108600;
  DFCid : UINT := 1231;
  debounceMethod : USINT := NATIVE;
END_STRUCT;
END_TYPE

TYPE DFC_SWReset : STRUCT
  DTC : UDINT := 16#105600;
  DFCid : UINT := 1308;
  debounceMethod : USINT := NATIVE;
END_STRUCT;
END_TYPE

TYPE DFC_MOXEMM_SMU_ALM2_23 : STRUCT
  DTC : UDINT := 16#108700;
  DFCid : UINT := 1232;
  debounceMethod : USINT := NATIVE;
END_STRUCT;
END_TYPE

TYPE DFC_MoXEMMHwLTMBIST : STRUCT
  DTC : UDINT := 16#10D100;
END_STRUCT;
END_TYPE

TYPE DFC_MOXEMM_SMU_ALM7_31 : STRUCT
  DTC : UDINT := 16#10B000;
  DFCid : UINT := 1278;
  debounceMethod : USINT := NATIVE;
END_STRUCT;
END_TYPE

TYPE DFC_MOXEMM_SMU_ALM7_30 : STRUCT
  DTC : UDINT := 16#10AF00;
  DFCid : UINT := 1277;
  debounceMethod : USINT := NATIVE;
END_STRUCT;
END_TYPE

TYPE DFC_OCWDAErrPin : STRUCT
  DTC : UDINT := 16#098B00;
  DFCid : UINT := 1307;
  debounceMethod : USINT := NATIVE;
END_STRUCT;
END_TYPE

TYPE DFC_ComCntESP_19 : STRUCT
  DTC : UDINT := 16#102500;
END_STRUCT;
END_TYPE

TYPE DFC_MOXEMM_SMU_ALM8_10 : STRUCT
  DTC : UDINT := 16#10B600;
  DFCid : UINT := 1281;
  debounceMethod : USINT := NATIVE;
END_STRUCT;
END_TYPE

TYPE DFC_MRlySCG : STRUCT
  DTC : UDINT := 16#104B00;
END_STRUCT;
END_TYPE

TYPE DFC_MOXEMM_SMU_ALM8_11 : STRUCT
  DTC : UDINT := 16#10B700;
  DFCid : UINT := 1282;
  debounceMethod : USINT := NATIVE;
END_STRUCT;
END_TYPE

TYPE DFC_MOXEMM_SMU_ALM8_12 : STRUCT
  DTC : UDINT := 16#10B800;
  DFCid : UINT := 1283;
  debounceMethod : USINT := NATIVE;
END_STRUCT;
END_TYPE

TYPE DFC_MOXEMM_SMU_ALM8_13 : STRUCT
  DTC : UDINT := 16#10B900;
  DFCid : UINT := 1284;
  debounceMethod : USINT := NATIVE;
END_STRUCT;
END_TYPE

TYPE DFC_MRlySCB : STRUCT
  DTC : UDINT := 16#104A00;
END_STRUCT;
END_TYPE

TYPE DFC_MoXEMMHwLTMCUFW : STRUCT
  DTC : UDINT := 16#10D200;
  DFCid : UINT := 1299;
  debounceMethod : USINT := NATIVE;
END_STRUCT;
END_TYPE

TYPE DFC_MOXEMM_SMU_ALM8_16 : STRUCT
  DTC : UDINT := 16#10BA00;
  DFCid : UINT := 1285;
  debounceMethod : USINT := NATIVE;
END_STRUCT;
END_TYPE

TYPE DFC_MOXEMM_SMU_ALM8_18 : STRUCT
  DTC : UDINT := 16#10BB00;
  DFCid : UINT := 1286;
  debounceMethod : USINT := NATIVE;
END_STRUCT;
END_TYPE

TYPE DFC_ComCntESP_10 : STRUCT
  DTC : UDINT := 16#102400;
END_STRUCT;
END_TYPE

TYPE DFC_CAN_E_TIMEOUT : STRUCT
  DTC : UDINT := 16#094200;
  DFCid : UINT := 1165;
  debounceMethod : USINT := NO_DEBOUNCE;
END_STRUCT;
END_TYPE

TYPE DFC_RBA_IOEXTLIB_KEEPALIVE_INI : STRUCT
  DTC : UDINT := 16#094400;
  DFCid : UINT := 1176;
  debounceMethod : USINT := NO_DEBOUNCE;
END_STRUCT;
END_TYPE

TYPE DFC_Com_vWhlRrL : STRUCT
  DTC : UDINT := 16#103D00;
END_STRUCT;
END_TYPE

TYPE DFC_Com_numWhlIncFrtLeft : STRUCT
  DTC : UDINT := 16#103A00;
END_STRUCT;
END_TYPE

TYPE DFC_rba_MemDiag_MemWrErr : STRUCT
  DTC : UDINT := 16#094800;
  DFCid : UINT := 1180;
  debounceMethod : USINT := NO_DEBOUNCE;
END_STRUCT;
END_TYPE

TYPE DFC_CANTRCV_E_NO_TRCV_CONTROL_0 : STRUCT
  DTC : UDINT := 16#094000;
  DFCid : UINT := 1164;
  debounceMethod : USINT := NO_DEBOUNCE;
END_STRUCT;
END_TYPE

TYPE DFC_MOXEMM_SMU_ALM3_11 : STRUCT
  DTC : UDINT := 16#108F00;
  DFCid : UINT := 1239;
  debounceMethod : USINT := NATIVE;
END_STRUCT;
END_TYPE

TYPE DFC_MOXEMM_SMU_ALM3_14 : STRUCT
  DTC : UDINT := 16#109100;
  DFCid : UINT := 1241;
  debounceMethod : USINT := NATIVE;
END_STRUCT;
END_TYPE

TYPE DFC_MOXEMM_SMU_ALM3_13 : STRUCT
  DTC : UDINT := 16#109000;
  DFCid : UINT := 1240;
  debounceMethod : USINT := NATIVE;
END_STRUCT;
END_TYPE

TYPE DFC_MOXEMM_SMU_ALM3_10 : STRUCT
  DTC : UDINT := 16#108E00;
  DFCid : UINT := 1238;
  debounceMethod : USINT := NATIVE;
END_STRUCT;
END_TYPE

TYPE DFC_MOXEMM_SMU_ALM8_30 : STRUCT
  DTC : UDINT := 16#10BC00;
  DFCid : UINT := 1289;
  debounceMethod : USINT := NATIVE;
END_STRUCT;
END_TYPE

TYPE DFC_MOXEMM_SMU_ALM8_31 : STRUCT
  DTC : UDINT := 16#10BD00;
  DFCid : UINT := 1290;
  debounceMethod : USINT := NATIVE;
END_STRUCT;
END_TYPE

TYPE DFC_ComCntACC_06 : STRUCT
  DTC : UDINT := 16#101F00;
END_STRUCT;
END_TYPE

TYPE DFC_rba_T15_Diag_ComInVld_Event : STRUCT
  DTC : UDINT := 16#094B00;
  DFCid : UINT := 1182;
  debounceMethod : USINT := NO_DEBOUNCE;
END_STRUCT;
END_TYPE

TYPE DFC_MOXEMM_SMU_ALM11_0 : STRUCT
  DTC : UDINT := 16#10C500;
  DFCid : UINT := 1201;
  debounceMethod : USINT := NATIVE;
END_STRUCT;
END_TYPE

TYPE DFC_MOXEMM_SMU_ALM11_1 : STRUCT
  DTC : UDINT := 16#10C600;
  DFCid : UINT := 1202;
  debounceMethod : USINT := NATIVE;
END_STRUCT;
END_TYPE

TYPE DFC_MOXEMM_SMU_ALM11_2 : STRUCT
  DTC : UDINT := 16#10C700;
  DFCid : UINT := 1203;
  debounceMethod : USINT := NATIVE;
END_STRUCT;
END_TYPE

TYPE DFC_MOXEMM_SMU_ALM3_23 : STRUCT
  DTC : UDINT := 16#109300;
  DFCid : UINT := 1244;
  debounceMethod : USINT := NATIVE;
END_STRUCT;
END_TYPE

TYPE DFC_MOXEMM_SMU_ALM3_22 : STRUCT
  DTC : UDINT := 16#109200;
  DFCid : UINT := 1243;
  debounceMethod : USINT := NATIVE;
END_STRUCT;
END_TYPE

TYPE DFC_OCWDACom : STRUCT
  DTC : UDINT := 16#098A00;
  DFCid : UINT := 1306;
  debounceMethod : USINT := NATIVE;
END_STRUCT;
END_TYPE

TYPE DFC_MoFVarPostBldSel : STRUCT
  DTC : UDINT := 16#098900;
  DFCid : UINT := 1297;
  debounceMethod : USINT := NATIVE;
END_STRUCT;
END_TYPE

TYPE DFC_MOXEMM_SMU_ALM1_2 : STRUCT
  DTC : UDINT := 16#107100;
  DFCid : UINT := 1215;
  debounceMethod : USINT := NATIVE;
END_STRUCT;
END_TYPE

TYPE DFC_MOXEMM_SMU_ALM1_4 : STRUCT
  DTC : UDINT := 16#107200;
  DFCid : UINT := 1218;
  debounceMethod : USINT := NATIVE;
END_STRUCT;
END_TYPE

TYPE DFC_MOXEMM_SMU_ALM1_5 : STRUCT
  DTC : UDINT := 16#107300;
  DFCid : UINT := 1219;
  debounceMethod : USINT := NATIVE;
END_STRUCT;
END_TYPE

TYPE DFC_MOXEMM_SMU_ALM1_7 : STRUCT
  DTC : UDINT := 16#107400;
  DFCid : UINT := 1220;
  debounceMethod : USINT := NATIVE;
END_STRUCT;
END_TYPE

TYPE DFC_MOXEMM_SMU_ALM1_8 : STRUCT
  DTC : UDINT := 16#107500;
  DFCid : UINT := 1221;
  debounceMethod : USINT := NATIVE;
END_STRUCT;
END_TYPE

TYPE DFC_MOXEMM_SMU_ALM9_0 : STRUCT
  DTC : UDINT := 16#10BE00;
  DFCid : UINT := 1292;
  debounceMethod : USINT := NATIVE;
END_STRUCT;
END_TYPE

TYPE DFC_MOXEMM_SMU_ALM9_1 : STRUCT
  DTC : UDINT := 16#10BF00;
  DFCid : UINT := 1293;
  debounceMethod : USINT := NATIVE;
END_STRUCT;
END_TYPE

TYPE DFC_ComChksBMS_01 : STRUCT
  DTC : UDINT := 16#101700;
END_STRUCT;
END_TYPE

TYPE DFC_LIN_E_TIMEOUT : STRUCT
  DTC : UDINT := 16#094100;
  DFCid : UINT := 1172;
  debounceMethod : USINT := NO_DEBOUNCE;
END_STRUCT;
END_TYPE

TYPE DFC_MOXEMM_SMU_ALM1_0 : STRUCT
  DTC : UDINT := 16#106F00;
  DFCid : UINT := 1209;
  debounceMethod : USINT := NATIVE;
END_STRUCT;
END_TYPE

TYPE DFC_MOXEMM_SMU_ALM1_1 : STRUCT
  DTC : UDINT := 16#107000;
  DFCid : UINT := 1210;
  debounceMethod : USINT := NATIVE;
END_STRUCT;
END_TYPE

TYPE DFC_MOXEMM_SMU_ALM1_14 : STRUCT
  DTC : UDINT := 16#107900;
  DFCid : UINT := 1214;
  debounceMethod : USINT := NATIVE;
END_STRUCT;
END_TYPE

TYPE DFC_MOXEMM_SMU_ALM1_13 : STRUCT
  DTC : UDINT := 16#107800;
  DFCid : UINT := 1213;
  debounceMethod : USINT := NATIVE;
END_STRUCT;
END_TYPE

TYPE DFC_MOXEMM_SMU_ALM1_10 : STRUCT
  DTC : UDINT := 16#107600;
  DFCid : UINT := 1211;
  debounceMethod : USINT := NATIVE;
END_STRUCT;
END_TYPE

TYPE DFC_rba_T15_Diag_ComOff_HwOn_Event : STRUCT
  DTC : UDINT := 16#094C00;
  DFCid : UINT := 1183;
  debounceMethod : USINT := NO_DEBOUNCE;
END_STRUCT;
END_TYPE

TYPE DFC_MOXEMM_SMU_ALM1_11 : STRUCT
  DTC : UDINT := 16#107700;
  DFCid : UINT := 1212;
  debounceMethod : USINT := NATIVE;
END_STRUCT;
END_TYPE

TYPE DFC_MOXEMM_SMU_ALM6_25 : STRUCT
  DTC : UDINT := 16#10A100;
  DFCid : UINT := 1259;
  debounceMethod : USINT := NATIVE;
END_STRUCT;
END_TYPE

TYPE DFC_MOXEMM_SMU_ALM6_21 : STRUCT
  DTC : UDINT := 16#10A000;
  DFCid : UINT := 1258;
  debounceMethod : USINT := NATIVE;
END_STRUCT;
END_TYPE

TYPE DFC_MOXEMM_SMU_ALM6_20 : STRUCT
  DTC : UDINT := 16#109F00;
  DFCid : UINT := 1257;
  debounceMethod : USINT := NATIVE;
END_STRUCT;
END_TYPE

TYPE DFC_ComDlcESP_02 : STRUCT
  DTC : UDINT := 16#102900;
END_STRUCT;
END_TYPE

TYPE DFC_MOXEMM_SMU_ALM1_23 : STRUCT
  DTC : UDINT := 16#107B00;
  DFCid : UINT := 1217;
  debounceMethod : USINT := NATIVE;
END_STRUCT;
END_TYPE

TYPE DFC_MOXEMM_SMU_ALM1_22 : STRUCT
  DTC : UDINT := 16#107A00;
  DFCid : UINT := 1216;
  debounceMethod : USINT := NATIVE;
END_STRUCT;
END_TYPE

TYPE DFC_rba_MRly_Diag_Stk_Event : STRUCT
  DTC : UDINT := 16#094600;
  DFCid : UINT := 1177;
  debounceMethod : USINT := NO_DEBOUNCE;
END_STRUCT;
END_TYPE

TYPE DFC_ComDlcESP_05 : STRUCT
  DTC : UDINT := 16#102A00;
END_STRUCT;
END_TYPE

TYPE DFC_DevLibBattULo : STRUCT
  DTC : UDINT := 16#092400;
  DFCid : UINT := 105;
  debounceMethod : USINT := TIME_UP_DOWN;
END_STRUCT;
END_TYPE

TYPE DFC_ComDlcESP_07 : STRUCT
  DTC : UDINT := 16#102B00;
END_STRUCT;
END_TYPE

TYPE DFC_MOXEMM_SMU_ALM2_1 : STRUCT
  DTC : UDINT := 16#107C00;
  DFCid : UINT := 1225;
  debounceMethod : USINT := NATIVE;
END_STRUCT;
END_TYPE

TYPE DFC_MOXEMM_SMU_ALM2_2 : STRUCT
  DTC : UDINT := 16#107D00;
  DFCid : UINT := 1230;
  debounceMethod : USINT := NATIVE;
END_STRUCT;
END_TYPE

TYPE DFC_MOXEMM_SMU_ALM2_4 : STRUCT
  DTC : UDINT := 16#107E00;
  DFCid : UINT := 1233;
  debounceMethod : USINT := NATIVE;
END_STRUCT;
END_TYPE

TYPE DFC_MOXEMM_SMU_ALM2_5 : STRUCT
  DTC : UDINT := 16#107F00;
  DFCid : UINT := 1234;
  debounceMethod : USINT := NATIVE;
END_STRUCT;
END_TYPE

TYPE DFC_MOXEMM_SMU_ALM2_7 : STRUCT
  DTC : UDINT := 16#108000;
  DFCid : UINT := 1235;
  debounceMethod : USINT := NATIVE;
END_STRUCT;
END_TYPE

TYPE DFC_MOXEMM_SMU_ALM2_8 : STRUCT
  DTC : UDINT := 16#108100;
  DFCid : UINT := 1236;
  debounceMethod : USINT := NATIVE;
END_STRUCT;
END_TYPE

TYPE DFC_rba_SyC_IrrSwOffTrigEngRun_Event : STRUCT
  DTC : UDINT := 16#094A00;
  DFCid : UINT := 1181;
  debounceMethod : USINT := NO_DEBOUNCE;
END_STRUCT;
END_TYPE

TYPE DFC_ComDlcESP_10 : STRUCT
  DTC : UDINT := 16#102C00;
END_STRUCT;
END_TYPE

TYPE DFC_MOXEMM_SMU_ALM7_17 : STRUCT
  DTC : UDINT := 16#10A900;
  DFCid : UINT := 1270;
  debounceMethod : USINT := NATIVE;
END_STRUCT;
END_TYPE

TYPE DFC_MOXEMM_SMU_ALM7_16 : STRUCT
  DTC : UDINT := 16#10A800;
  DFCid : UINT := 1269;
  debounceMethod : USINT := NATIVE;
END_STRUCT;
END_TYPE

TYPE DFC_MOXEMM_SMU_ALM7_15 : STRUCT
  DTC : UDINT := 16#10A700;
  DFCid : UINT := 1268;
  debounceMethod : USINT := NATIVE;
END_STRUCT;
END_TYPE

TYPE DFC_MOXEMM_SMU_ALM7_14 : STRUCT
  DTC : UDINT := 16#10A600;
  DFCid : UINT := 1267;
  debounceMethod : USINT := NATIVE;
END_STRUCT;
END_TYPE

TYPE DFC_MOXEMM_SMU_ALM7_13 : STRUCT
  DTC : UDINT := 16#10A500;
  DFCid : UINT := 1266;
  debounceMethod : USINT := NATIVE;
END_STRUCT;
END_TYPE

TYPE DFC_MOXEMM_SMU_ALM7_12 : STRUCT
  DTC : UDINT := 16#10A400;
  DFCid : UINT := 1265;
  debounceMethod : USINT := NATIVE;
END_STRUCT;
END_TYPE

TYPE DFC_ComDlcESP_19 : STRUCT
  DTC : UDINT := 16#102D00;
END_STRUCT;
END_TYPE

TYPE DFC_ComCntKlemmen_Status_01 : STRUCT
  DTC : UDINT := 16#103900;
END_STRUCT;
END_TYPE

TYPE DFC_rba_T15_Diag_ComOn_HwOff_Event : STRUCT
  DTC : UDINT := 16#094D00;
  DFCid : UINT := 1184;
  debounceMethod : USINT := NO_DEBOUNCE;
END_STRUCT;
END_TYPE

TYPE DFC_MoXEMMHwLTStbySMUAlvTest : STRUCT
  DTC : UDINT := 16#10D500;
  DFCid : UINT := 1302;
  debounceMethod : USINT := NATIVE;
END_STRUCT;
END_TYPE

TYPE DFC_rba_MultiStackTrace_Threshold : STRUCT
  DTC : UDINT := 16#094900;
  DFCid : UINT := 1173;
  debounceMethod : USINT := NO_DEBOUNCE;
END_STRUCT;
END_TYPE

TYPE DFC_MOXEMM_SMU_ALM2_14 : STRUCT
  DTC : UDINT := 16#108500;
  DFCid : UINT := 1229;
  debounceMethod : USINT := NATIVE;
END_STRUCT;
END_TYPE

TYPE DFC_ComDlcESP_20 : STRUCT
  DTC : UDINT := 16#102E00;
END_STRUCT;
END_TYPE

TYPE DFC_MOXEMM_SMU_ALM2_11 : STRUCT
  DTC : UDINT := 16#108300;
  DFCid : UINT := 1227;
  debounceMethod : USINT := NATIVE;
END_STRUCT;
END_TYPE

TYPE DFC_MOXEMM_SMU_ALM7_29 : STRUCT
  DTC : UDINT := 16#10AE00;
  DFCid : UINT := 1276;
  debounceMethod : USINT := NATIVE;
END_STRUCT;
END_TYPE

TYPE DFC_ComDlcESP_21 : STRUCT
  DTC : UDINT := 16#102F00;
END_STRUCT;
END_TYPE

TYPE DFC_MOXEMM_SMU_ALM2_10 : STRUCT
  DTC : UDINT := 16#108200;
  DFCid : UINT := 1226;
  debounceMethod : USINT := NATIVE;
END_STRUCT;
END_TYPE

TYPE DFC_MOXEMM_SMU_ALM7_28 : STRUCT
  DTC : UDINT := 16#10AD00;
  DFCid : UINT := 1275;
  debounceMethod : USINT := NATIVE;
END_STRUCT;
END_TYPE

TYPE DFC_MOXEMM_SMU_ALM2_13 : STRUCT
  DTC : UDINT := 16#108400;
  DFCid : UINT := 1228;
  debounceMethod : USINT := NATIVE;
END_STRUCT;
END_TYPE

TYPE DFC_MOXEMM_SMU_ALM7_26 : STRUCT
  DTC : UDINT := 16#10AC00;
  DFCid : UINT := 1274;
  debounceMethod : USINT := NATIVE;
END_STRUCT;
END_TYPE

TYPE DFC_MOXEMM_SMU_ALM3_8 : STRUCT
  DTC : UDINT := 16#108D00;
  DFCid : UINT := 1248;
  debounceMethod : USINT := NATIVE;
END_STRUCT;
END_TYPE

TYPE DFC_MOXEMM_SMU_ALM7_25 : STRUCT
  DTC : UDINT := 16#10AB00;
  DFCid : UINT := 1273;
  debounceMethod : USINT := NATIVE;
END_STRUCT;
END_TYPE

TYPE DFC_MOXEMM_SMU_ALM7_20 : STRUCT
  DTC : UDINT := 16#10AA00;
  DFCid : UINT := 1272;
  debounceMethod : USINT := NATIVE;
END_STRUCT;
END_TYPE

TYPE DFC_MRlyOL : STRUCT
  DTC : UDINT := 16#104900;
END_STRUCT;
END_TYPE

TYPE DFC_MOXEMM_SMU_ALM7_1 : STRUCT
  DTC : UDINT := 16#10A200;
  DFCid : UINT := 1264;
  debounceMethod : USINT := NATIVE;
END_STRUCT;
END_TYPE

TYPE DFC_ComChksESP_19 : STRUCT
  DTC : UDINT := 16#101C00;
END_STRUCT;
END_TYPE

TYPE DFC_MOXEMM_SMU_ALM7_2 : STRUCT
  DTC : UDINT := 16#10A300;
  DFCid : UINT := 1271;
  debounceMethod : USINT := NATIVE;
END_STRUCT;
END_TYPE

TYPE DFC_ComTOutESP_10 : STRUCT
  DTC : UDINT := 16#103400;
END_STRUCT;
END_TYPE

TYPE DFC_Com_stWhlSensRrRht : STRUCT
  DTC : UDINT := 16#103B00;
END_STRUCT;
END_TYPE

TYPE DFC_ComChksKlemmen_Status_01 : STRUCT
  DTC : UDINT := 16#103800;
END_STRUCT;
END_TYPE

TYPE DFC_ComTOutESP_07 : STRUCT
  DTC : UDINT := 16#103300;
END_STRUCT;
END_TYPE

TYPE DFC_ComDlcACC_06 : STRUCT
  DTC : UDINT := 16#102800;
END_STRUCT;
END_TYPE

TYPE DFC_rba_MemDiag_MemReadErr : STRUCT
  DTC : UDINT := 16#094700;
  DFCid : UINT := 1179;
  debounceMethod : USINT := NO_DEBOUNCE;
END_STRUCT;
END_TYPE

TYPE DFC_ComChksESP_10 : STRUCT
  DTC : UDINT := 16#101B00;
END_STRUCT;
END_TYPE

TYPE DFC_ComChksESP_05 : STRUCT
  DTC : UDINT := 16#101900;
END_STRUCT;
END_TYPE

TYPE DFC_OCWDAABEActv : STRUCT
  DTC : UDINT := 16#10D800;
  DFCid : UINT := 1305;
  debounceMethod : USINT := NATIVE;
END_STRUCT;
END_TYPE

TYPE DFC_ComChksESP_07 : STRUCT
  DTC : UDINT := 16#101A00;
END_STRUCT;
END_TYPE

TYPE DFC_ComTOutESP_21 : STRUCT
  DTC : UDINT := 16#103700;
END_STRUCT;
END_TYPE

TYPE DFC_ComTOutESP_20 : STRUCT
  DTC : UDINT := 16#103600;
END_STRUCT;
END_TYPE

TYPE DFC_MOXEMM_SMU_ALM0_13 : STRUCT
  DTC : UDINT := 16#106B00;
  DFCid : UINT := 1189;
  debounceMethod : USINT := NATIVE;
END_STRUCT;
END_TYPE

TYPE DFC_MOXEMM_SMU_ALM0_14 : STRUCT
  DTC : UDINT := 16#106C00;
  DFCid : UINT := 1190;
  debounceMethod : USINT := NATIVE;
END_STRUCT;
END_TYPE

TYPE DFC_ComTOutESP_19 : STRUCT
  DTC : UDINT := 16#103500;
END_STRUCT;
END_TYPE

TYPE DFC_MOXEMM_SMU_ALM0_10 : STRUCT
  DTC : UDINT := 16#106900;
  DFCid : UINT := 1187;
  debounceMethod : USINT := NATIVE;
END_STRUCT;
END_TYPE

TYPE DFC_MOXEMM_SMU_ALM0_11 : STRUCT
  DTC : UDINT := 16#106A00;
  DFCid : UINT := 1188;
  debounceMethod : USINT := NATIVE;
END_STRUCT;
END_TYPE

TYPE DFC_MOXEMM_SMU_ALM8_3 : STRUCT
  DTC : UDINT := 16#10B400;
  DFCid : UINT := 1288;
  debounceMethod : USINT := NATIVE;
END_STRUCT;
END_TYPE

TYPE DFC_MOXEMM_SMU_ALM8_4 : STRUCT
  DTC : UDINT := 16#10B500;
  DFCid : UINT := 1291;
  debounceMethod : USINT := NATIVE;
END_STRUCT;
END_TYPE

TYPE DFC_ComChksESP_02 : STRUCT
  DTC : UDINT := 16#101800;
END_STRUCT;
END_TYPE

TYPE DFC_DevLibBattUHi : STRUCT
  DTC : UDINT := 16#092300;
  DFCid : UINT := 104;
  debounceMethod : USINT := TIME_UP_DOWN;
END_STRUCT;
END_TYPE

TYPE DFC_Com_trqClthTCSDCSDes : STRUCT
  DTC : UDINT := 16#103C00;
END_STRUCT;
END_TYPE

TYPE DFC_MOXEMM_SMU_ALM0_4 : STRUCT
  DTC : UDINT := 16#106500;
  DFCid : UINT := 1194;
  debounceMethod : USINT := NATIVE;
END_STRUCT;
END_TYPE

TYPE DFC_MoXEMMHwLTTempSens : STRUCT
  DTC : UDINT := 16#10D600;
  DFCid : UINT := 1303;
  debounceMethod : USINT := NATIVE;
END_STRUCT;
END_TYPE

TYPE DFC_MOXEMM_SMU_ALM0_5 : STRUCT
  DTC : UDINT := 16#106600;
  DFCid : UINT := 1195;
  debounceMethod : USINT := NATIVE;
END_STRUCT;
END_TYPE

TYPE DFC_MOXEMM_SMU_ALM0_7 : STRUCT
  DTC : UDINT := 16#106700;
  DFCid : UINT := 1196;
  debounceMethod : USINT := NATIVE;
END_STRUCT;
END_TYPE

TYPE DFC_MOXEMM_SMU_ALM0_8 : STRUCT
  DTC : UDINT := 16#106800;
  DFCid : UINT := 1197;
  debounceMethod : USINT := NATIVE;
END_STRUCT;
END_TYPE

TYPE DFC_MOXEMM_SMU_ALM8_0 : STRUCT
  DTC : UDINT := 16#10B100;
  DFCid : UINT := 1279;
  debounceMethod : USINT := NATIVE;
END_STRUCT;
END_TYPE

TYPE DFC_MOXEMM_SMU_ALM8_1 : STRUCT
  DTC : UDINT := 16#10B200;
  DFCid : UINT := 1280;
  debounceMethod : USINT := NATIVE;
END_STRUCT;
END_TYPE

TYPE DFC_MOXEMM_SMU_ALM8_2 : STRUCT
  DTC : UDINT := 16#10B300;
  DFCid : UINT := 1287;
  debounceMethod : USINT := NATIVE;
END_STRUCT;
END_TYPE

TYPE DFC_ComChksACC_06 : STRUCT
  DTC : UDINT := 16#101600;
END_STRUCT;
END_TYPE

TYPE DFC_MOXEMM_SMU_ALM0_0 : STRUCT
  DTC : UDINT := 16#106200;
  DFCid : UINT := 1185;
  debounceMethod : USINT := NATIVE;
END_STRUCT;
END_TYPE

TYPE DFC_MOXEMM_SMU_ALM0_1 : STRUCT
  DTC : UDINT := 16#106300;
  DFCid : UINT := 1186;
  debounceMethod : USINT := NATIVE;
END_STRUCT;
END_TYPE

TYPE DFC_SWReset_2 : STRUCT
  DTC : UDINT := 16#105900;
END_STRUCT;
END_TYPE

TYPE DFC_MOXEMM_SMU_ALM0_2 : STRUCT
  DTC : UDINT := 16#106400;
  DFCid : UINT := 1191;
  debounceMethod : USINT := NATIVE;
END_STRUCT;
END_TYPE

TYPE DFC_MOXEMM_SMU_ALM0_23 : STRUCT
  DTC : UDINT := 16#106E00;
  DFCid : UINT := 1193;
  debounceMethod : USINT := NATIVE;
END_STRUCT;
END_TYPE

TYPE DFC_MOXEMM_SMU_ALM0_22 : STRUCT
  DTC : UDINT := 16#106D00;
  DFCid : UINT := 1192;
  debounceMethod : USINT := NATIVE;
END_STRUCT;
END_TYPE

TYPE DFC_ComTOutESP_05 : STRUCT
  DTC : UDINT := 16#103200;
END_STRUCT;
END_TYPE

TYPE DFC_ComTOutESP_02 : STRUCT
  DTC : UDINT := 16#103100;
END_STRUCT;
END_TYPE

TYPE DFC_MOXEMM_SMU_ALM6_18 : STRUCT
  DTC : UDINT := 16#109E00;
  DFCid : UINT := 1255;
  debounceMethod : USINT := NATIVE;
END_STRUCT;
END_TYPE

TYPE DFC_MOXEMM_SMU_ALM6_17 : STRUCT
  DTC : UDINT := 16#109D00;
  DFCid : UINT := 1254;
  debounceMethod : USINT := NATIVE;
END_STRUCT;
END_TYPE

TYPE DFC_MOXEMM_SMU_ALM6_15 : STRUCT
  DTC : UDINT := 16#109C00;
  DFCid : UINT := 1253;
  debounceMethod : USINT := NATIVE;
END_STRUCT;
END_TYPE

TYPE DFC_MOXEMM_SMU_ALM21_16 : STRUCT
  DTC : UDINT := 16#10CF00;
  DFCid : UINT := 1223;
  debounceMethod : USINT := NATIVE;
END_STRUCT;
END_TYPE

TYPE DFC_MOXEMM_SMU_ALM6_14 : STRUCT
  DTC : UDINT := 16#109B00;
  DFCid : UINT := 1252;
  debounceMethod : USINT := NATIVE;
END_STRUCT;
END_TYPE

TYPE DFC_MOXEMM_SMU_ALM6_12 : STRUCT
  DTC : UDINT := 16#109A00;
  DFCid : UINT := 1251;
  debounceMethod : USINT := NATIVE;
END_STRUCT;
END_TYPE

TYPE DFC_MOXEMM_SMU_ALM9_3 : STRUCT
  DTC : UDINT := 16#10C000;
  DFCid : UINT := 1295;
  debounceMethod : USINT := NATIVE;
END_STRUCT;
END_TYPE

TYPE DFC_MOXEMM_SMU_ALM6_11 : STRUCT
  DTC : UDINT := 16#109900;
  DFCid : UINT := 1250;
  debounceMethod : USINT := NATIVE;
END_STRUCT;
END_TYPE

TYPE DFC_ComTOutACC_06 : STRUCT
  DTC : UDINT := 16#103000;
END_STRUCT;
END_TYPE

TYPE DFC_MOXEMM_SMU_ALM9_15 : STRUCT
  DTC : UDINT := 16#10C100;
  DFCid : UINT := 1294;
  debounceMethod : USINT := NATIVE;
END_STRUCT;
END_TYPE

TYPE DFC_MOXEMM_SMU_ALM11_8 : STRUCT
  DTC : UDINT := 16#10CB00;
  DFCid : UINT := 1207;
  debounceMethod : USINT := NATIVE;
END_STRUCT;
END_TYPE

TYPE DFC_MOXEMM_SMU_ALM11_9 : STRUCT
  DTC : UDINT := 16#10CC00;
  DFCid : UINT := 1208;
  debounceMethod : USINT := NATIVE;
END_STRUCT;
END_TYPE

TYPE DFC_MOXEMM_SMU_ALM11_3 : STRUCT
  DTC : UDINT := 16#10C800;
  DFCid : UINT := 1204;
  debounceMethod : USINT := NATIVE;
END_STRUCT;
END_TYPE

TYPE DFC_MOXEMM_SMU_ALM11_4 : STRUCT
  DTC : UDINT := 16#10C900;
  DFCid : UINT := 1205;
  debounceMethod : USINT := NATIVE;
END_STRUCT;
END_TYPE

TYPE DFC_MOXEMM_SMU_ALM11_5 : STRUCT
  DTC : UDINT := 16#10CA00;
  DFCid : UINT := 1206;
  debounceMethod : USINT := NATIVE;
END_STRUCT;
END_TYPE

TYPE DFC_MOXEMM_SMU_ALM10_16 : STRUCT
  DTC : UDINT := 16#10C200;
  DFCid : UINT := 1198;
  debounceMethod : USINT := NATIVE;
END_STRUCT;
END_TYPE

TYPE DFC_MOXEMM_SMU_ALM10_17 : STRUCT
  DTC : UDINT := 16#10C300;
  DFCid : UINT := 1199;
  debounceMethod : USINT := NATIVE;
END_STRUCT;
END_TYPE

TYPE DFC_MoXEMMHwLTUCBCfg : STRUCT
  DTC : UDINT := 16#10D700;
  DFCid : UINT := 1304;
  debounceMethod : USINT := NATIVE;
END_STRUCT;
END_TYPE

TYPE DFC_CANSM_E_BUS_OFF_NETWORK_0 : STRUCT
  DTC : UDINT := 16#104C00;
  DFCid : UINT := 1160;
  debounceMethod : USINT := NO_DEBOUNCE;
END_STRUCT;
END_TYPE

TYPE DFC_CANSM_E_BUS_OFF_NETWORK_3 : STRUCT
  DTC : UDINT := 16#104F00;
  DFCid : UINT := 1163;
  debounceMethod : USINT := NO_DEBOUNCE;
END_STRUCT;
END_TYPE

TYPE DFC_CANSM_E_BUS_OFF_NETWORK_1 : STRUCT
  DTC : UDINT := 16#104D00;
  DFCid : UINT := 1161;
  debounceMethod : USINT := NO_DEBOUNCE;
END_STRUCT;
END_TYPE

TYPE DFC_CANSM_E_BUS_OFF_NETWORK_2 : STRUCT
  DTC : UDINT := 16#104E00;
  DFCid : UINT := 1162;
  debounceMethod : USINT := NO_DEBOUNCE;
END_STRUCT;
END_TYPE

TYPE DFC_ComCntBMS_01 : STRUCT
  DTC : UDINT := 16#102000;
END_STRUCT;
END_TYPE

TYPE DFC_MoXEMMHwLTLBIST : STRUCT
  DTC : UDINT := 16#10D000;
END_STRUCT;
END_TYPE

TYPE DFC_MoXEMMHwLTMonBIST : STRUCT
  DTC : UDINT := 16#10D300;
  DFCid : UINT := 1300;
  debounceMethod : USINT := NATIVE;
END_STRUCT;
END_TYPE

TYPE DFC_SWReset_1 : STRUCT
  DTC : UDINT := 16#105800;
END_STRUCT;
END_TYPE

TYPE DFC_SWReset_0 : STRUCT
  DTC : UDINT := 16#105700;
END_STRUCT;
END_TYPE

TYPE DFC_rba_MemDiagExtd_MemReadSngErr : STRUCT
  DTC : UDINT := 16#103E00;
  DFCid : UINT := 1178;
  debounceMethod : USINT := NO_DEBOUNCE;
END_STRUCT;
END_TYPE

TYPE DFC_MOXEMM_SMU_ALM10_21 : STRUCT
  DTC : UDINT := 16#10C400;
  DFCid : UINT := 1200;
  debounceMethod : USINT := NATIVE;
END_STRUCT;
END_TYPE

TYPE DFC_MOXEMM_SMU_ALM6_5 : STRUCT
  DTC : UDINT := 16#109600;
  DFCid : UINT := 1261;
  debounceMethod : USINT := NATIVE;
END_STRUCT;
END_TYPE

TYPE DFC_MOXEMM_SMU_ALM6_7 : STRUCT
  DTC : UDINT := 16#109700;
  DFCid : UINT := 1262;
  debounceMethod : USINT := NATIVE;
END_STRUCT;
END_TYPE

TYPE DFC_MOXEMM_SMU_ALM6_8 : STRUCT
  DTC : UDINT := 16#109800;
  DFCid : UINT := 1263;
  debounceMethod : USINT := NATIVE;
END_STRUCT;
END_TYPE

TYPE DFC_COMM_E_NET_START_IND_CHANNEL_3 : STRUCT
  DTC : UDINT := 16#105300;
  DFCid : UINT := 1169;
  debounceMethod : USINT := NO_DEBOUNCE;
END_STRUCT;
END_TYPE

TYPE DFC_COMM_E_NET_START_IND_CHANNEL_2 : STRUCT
  DTC : UDINT := 16#105200;
  DFCid : UINT := 1168;
  debounceMethod : USINT := NO_DEBOUNCE;
END_STRUCT;
END_TYPE

TYPE DFC_COMM_E_NET_START_IND_CHANNEL_5 : STRUCT
  DTC : UDINT := 16#105500;
  DFCid : UINT := 1171;
  debounceMethod : USINT := NO_DEBOUNCE;
END_STRUCT;
END_TYPE

TYPE DFC_COMM_E_NET_START_IND_CHANNEL_4 : STRUCT
  DTC : UDINT := 16#105400;
  DFCid : UINT := 1170;
  debounceMethod : USINT := NO_DEBOUNCE;
END_STRUCT;
END_TYPE

TYPE DFC_MOXEMM_SMU_ALM6_0 : STRUCT
  DTC : UDINT := 16#109400;
  DFCid : UINT := 1249;
  debounceMethod : USINT := NATIVE;
END_STRUCT;
END_TYPE

TYPE DFC_MOXEMM_SMU_ALM6_2 : STRUCT
  DTC : UDINT := 16#10D900;
  DFCid : UINT := 1256;
  debounceMethod : USINT := NATIVE;
END_STRUCT;
END_TYPE

TYPE DFC_MOXEMM_SMU_ALM6_4 : STRUCT
  DTC : UDINT := 16#109500;
  DFCid : UINT := 1260;
  debounceMethod : USINT := NATIVE;
END_STRUCT;
END_TYPE

TYPE DFC_ComCntESP_20 : STRUCT
  DTC : UDINT := 16#102600;
END_STRUCT;
END_TYPE

TYPE DFC_ComCntESP_21 : STRUCT
  DTC : UDINT := 16#102700;
END_STRUCT;
END_TYPE

TYPE DFC_COMM_E_NET_START_IND_CHANNEL_1 : STRUCT
  DTC : UDINT := 16#105100;
  DFCid : UINT := 1167;
  debounceMethod : USINT := NO_DEBOUNCE;
END_STRUCT;
END_TYPE

TYPE DFC_COMM_E_NET_START_IND_CHANNEL_0 : STRUCT
  DTC : UDINT := 16#105000;
  DFCid : UINT := 1166;
  debounceMethod : USINT := NO_DEBOUNCE;
END_STRUCT;
END_TYPE

TYPE DFC_MOXEMM_SMU_ALM21_0 : STRUCT
  DTC : UDINT := 16#10CD00;
  DFCid : UINT := 1222;
  debounceMethod : USINT := NATIVE;
END_STRUCT;
END_TYPE

TYPE DFC_MoCSOPICO : STRUCT
  DTC : UDINT := 16#106000;
  DFCid : UINT := 1296;
  debounceMethod : USINT := NATIVE;
END_STRUCT;
END_TYPE

TYPE DFC_MOXEMM_SMU_ALM21_3 : STRUCT
  DTC : UDINT := 16#10CE00;
  DFCid : UINT := 1224;
  debounceMethod : USINT := NATIVE;
END_STRUCT;
END_TYPE

TYPE DFC_MoSysCtrlReIni : STRUCT
  DTC : UDINT := 16#106100;
  DFCid : UINT := 1298;
  debounceMethod : USINT := NATIVE;
END_STRUCT;
END_TYPE

TYPE DFC_RBA_IOEXTLIB_KEEPALIVE_DRV : STRUCT
  DTC : UDINT := 16#094300;
  DFCid : UINT := 1175;
  debounceMethod : USINT := NO_DEBOUNCE;
END_STRUCT;
END_TYPE

TYPE DFC_ComChksESP_20 : STRUCT
  DTC : UDINT := 16#101D00;
END_STRUCT;
END_TYPE

TYPE DFC_ComChksESP_21 : STRUCT
  DTC : UDINT := 16#101E00;
END_STRUCT;
END_TYPE

TYPE DFC_bds_TiUpDwn0x8A01 : STRUCT
  DTC : UDINT := 16#8A0100;
  DFCid : UINT := 206;
  debounceMethod : USINT := TIME_UP_DOWN;
END_STRUCT;
END_TYPE

TYPE DFC_bds_TiUpDwn0x8A02 : STRUCT
  DTC : UDINT := 16#8A0200;
  DFCid : UINT := 207;
  debounceMethod : USINT := TIME_UP_DOWN;
END_STRUCT;
END_TYPE

TYPE DFC_bds_TiUpDwn0x8A03 : STRUCT
  DTC : UDINT := 16#8A0300;
  DFCid : UINT := 208;
  debounceMethod : USINT := TIME_UP_DOWN;
END_STRUCT;
END_TYPE

TYPE DFC_bds_TiInRow0x8B01 : STRUCT
  DTC : UDINT := 16#8B0100;
  DFCid : UINT := 101;
  debounceMethod : USINT := TIME_IN_ROW;
END_STRUCT;
END_TYPE

TYPE DFC_bds_TiInRow0x8B02 : STRUCT
  DTC : UDINT := 16#8B0200;
  DFCid : UINT := 102;
  debounceMethod : USINT := TIME_IN_ROW;
END_STRUCT;
END_TYPE

TYPE DFC_bds_TiInRow0x8B03 : STRUCT
  DTC : UDINT := 16#8B0300;
  DFCid : UINT := 103;
  debounceMethod : USINT := TIME_IN_ROW;
END_STRUCT;
END_TYPE

TYPE DFC_bds_NoDeb0x8C01 : STRUCT
  DTC : UDINT := 16#8C0100;
  DFCid : UINT := 820;
  debounceMethod : USINT := NO_DEBOUNCE;
END_STRUCT;
END_TYPE

TYPE DFC_bds_NoDeb0x8C02 : STRUCT
  DTC : UDINT := 16#8C0200;
  DFCid : UINT := 821;
  debounceMethod : USINT := NO_DEBOUNCE;
END_STRUCT;
END_TYPE

TYPE DFC_bds_NoDeb0x8C03 : STRUCT
  DTC : UDINT := 16#8C0300;
  DFCid : UINT := 822;
  debounceMethod : USINT := NO_DEBOUNCE;
END_STRUCT;
END_TYPE

TYPE DFC_bds_NoDeb0x8000 : STRUCT
  DTC : UDINT := 16#800000;
  DFCid : UINT := 721;
  debounceMethod : USINT := NO_DEBOUNCE;
END_STRUCT;
END_TYPE

TYPE DFC_bds_NoDeb0x8001 : STRUCT
  DTC : UDINT := 16#800100;
  DFCid : UINT := 722;
  debounceMethod : USINT := NO_DEBOUNCE;
END_STRUCT;
END_TYPE

TYPE DFC_bds_NoDeb0x8002 : STRUCT
  DTC : UDINT := 16#800200;
  DFCid : UINT := 723;
  debounceMethod : USINT := NO_DEBOUNCE;
END_STRUCT;
END_TYPE

TYPE DFC_bds_NoDeb0x8003 : STRUCT
  DTC : UDINT := 16#800300;
  DFCid : UINT := 724;
  debounceMethod : USINT := NO_DEBOUNCE;
END_STRUCT;
END_TYPE

TYPE DFC_bds_NoDeb0x8004 : STRUCT
  DTC : UDINT := 16#800400;
  DFCid : UINT := 725;
  debounceMethod : USINT := NO_DEBOUNCE;
END_STRUCT;
END_TYPE

TYPE DFC_bds_NoDeb0x8005 : STRUCT
  DTC : UDINT := 16#800500;
  DFCid : UINT := 726;
  debounceMethod : USINT := NO_DEBOUNCE;
END_STRUCT;
END_TYPE

TYPE DFC_bds_NoDeb0x8006 : STRUCT
  DTC : UDINT := 16#800600;
  DFCid : UINT := 727;
  debounceMethod : USINT := NO_DEBOUNCE;
END_STRUCT;
END_TYPE

TYPE DFC_bds_NoDeb0x8007 : STRUCT
  DTC : UDINT := 16#800700;
  DFCid : UINT := 728;
  debounceMethod : USINT := NO_DEBOUNCE;
END_STRUCT;
END_TYPE

TYPE DFC_bds_NoDeb0x8008 : STRUCT
  DTC : UDINT := 16#800800;
  DFCid : UINT := 729;
  debounceMethod : USINT := NO_DEBOUNCE;
END_STRUCT;
END_TYPE

TYPE DFC_bds_NoDeb0x8009 : STRUCT
  DTC : UDINT := 16#800900;
  DFCid : UINT := 730;
  debounceMethod : USINT := NO_DEBOUNCE;
END_STRUCT;
END_TYPE

TYPE DFC_bds_NoDeb0x800a : STRUCT
  DTC : UDINT := 16#800A00;
  DFCid : UINT := 731;
  debounceMethod : USINT := NO_DEBOUNCE;
END_STRUCT;
END_TYPE

TYPE DFC_bds_NoDeb0x800b : STRUCT
  DTC : UDINT := 16#800B00;
  DFCid : UINT := 732;
  debounceMethod : USINT := NO_DEBOUNCE;
END_STRUCT;
END_TYPE

TYPE DFC_bds_NoDeb0x800c : STRUCT
  DTC : UDINT := 16#800C00;
  DFCid : UINT := 733;
  debounceMethod : USINT := NO_DEBOUNCE;
END_STRUCT;
END_TYPE

TYPE DFC_bds_NoDeb0x800d : STRUCT
  DTC : UDINT := 16#800D00;
  DFCid : UINT := 734;
  debounceMethod : USINT := NO_DEBOUNCE;
END_STRUCT;
END_TYPE

TYPE DFC_bds_NoDeb0x800e : STRUCT
  DTC : UDINT := 16#800E00;
  DFCid : UINT := 735;
  debounceMethod : USINT := NO_DEBOUNCE;
END_STRUCT;
END_TYPE

TYPE DFC_bds_NoDeb0x800f : STRUCT
  DTC : UDINT := 16#800F00;
  DFCid : UINT := 736;
  debounceMethod : USINT := NO_DEBOUNCE;
END_STRUCT;
END_TYPE

TYPE DFC_bds_NoDeb0x8010 : STRUCT
  DTC : UDINT := 16#801000;
  DFCid : UINT := 737;
  debounceMethod : USINT := NO_DEBOUNCE;
END_STRUCT;
END_TYPE

TYPE DFC_bds_NoDeb0x8011 : STRUCT
  DTC : UDINT := 16#801100;
  DFCid : UINT := 738;
  debounceMethod : USINT := NO_DEBOUNCE;
END_STRUCT;
END_TYPE

TYPE DFC_bds_NoDeb0x8012 : STRUCT
  DTC : UDINT := 16#801200;
  DFCid : UINT := 739;
  debounceMethod : USINT := NO_DEBOUNCE;
END_STRUCT;
END_TYPE

TYPE DFC_bds_NoDeb0x8013 : STRUCT
  DTC : UDINT := 16#801300;
  DFCid : UINT := 740;
  debounceMethod : USINT := NO_DEBOUNCE;
END_STRUCT;
END_TYPE

TYPE DFC_bds_NoDeb0x8014 : STRUCT
  DTC : UDINT := 16#801400;
  DFCid : UINT := 741;
  debounceMethod : USINT := NO_DEBOUNCE;
END_STRUCT;
END_TYPE

TYPE DFC_bds_NoDeb0x8015 : STRUCT
  DTC : UDINT := 16#801500;
  DFCid : UINT := 742;
  debounceMethod : USINT := NO_DEBOUNCE;
END_STRUCT;
END_TYPE

TYPE DFC_bds_NoDeb0x8016 : STRUCT
  DTC : UDINT := 16#801600;
  DFCid : UINT := 743;
  debounceMethod : USINT := NO_DEBOUNCE;
END_STRUCT;
END_TYPE

TYPE DFC_bds_NoDeb0x8017 : STRUCT
  DTC : UDINT := 16#801700;
  DFCid : UINT := 744;
  debounceMethod : USINT := NO_DEBOUNCE;
END_STRUCT;
END_TYPE

TYPE DFC_bds_NoDeb0x8018 : STRUCT
  DTC : UDINT := 16#801800;
  DFCid : UINT := 745;
  debounceMethod : USINT := NO_DEBOUNCE;
END_STRUCT;
END_TYPE

TYPE DFC_bds_NoDeb0x8019 : STRUCT
  DTC : UDINT := 16#801900;
  DFCid : UINT := 746;
  debounceMethod : USINT := NO_DEBOUNCE;
END_STRUCT;
END_TYPE

TYPE DFC_bds_NoDeb0x801a : STRUCT
  DTC : UDINT := 16#801A00;
  DFCid : UINT := 747;
  debounceMethod : USINT := NO_DEBOUNCE;
END_STRUCT;
END_TYPE

TYPE DFC_bds_NoDeb0x801b : STRUCT
  DTC : UDINT := 16#801B00;
  DFCid : UINT := 748;
  debounceMethod : USINT := NO_DEBOUNCE;
END_STRUCT;
END_TYPE

TYPE DFC_bds_NoDeb0x801c : STRUCT
  DTC : UDINT := 16#801C00;
  DFCid : UINT := 749;
  debounceMethod : USINT := NO_DEBOUNCE;
END_STRUCT;
END_TYPE

TYPE DFC_bds_NoDeb0x801d : STRUCT
  DTC : UDINT := 16#801D00;
  DFCid : UINT := 750;
  debounceMethod : USINT := NO_DEBOUNCE;
END_STRUCT;
END_TYPE

TYPE DFC_bds_NoDeb0x801e : STRUCT
  DTC : UDINT := 16#801E00;
  DFCid : UINT := 751;
  debounceMethod : USINT := NO_DEBOUNCE;
END_STRUCT;
END_TYPE

TYPE DFC_bds_NoDeb0x801f : STRUCT
  DTC : UDINT := 16#801F00;
  DFCid : UINT := 752;
  debounceMethod : USINT := NO_DEBOUNCE;
END_STRUCT;
END_TYPE

TYPE DFC_bds_NoDeb0x8020 : STRUCT
  DTC : UDINT := 16#802000;
  DFCid : UINT := 753;
  debounceMethod : USINT := NO_DEBOUNCE;
END_STRUCT;
END_TYPE

TYPE DFC_bds_NoDeb0x8021 : STRUCT
  DTC : UDINT := 16#802100;
  DFCid : UINT := 754;
  debounceMethod : USINT := NO_DEBOUNCE;
END_STRUCT;
END_TYPE

TYPE DFC_bds_NoDeb0x8022 : STRUCT
  DTC : UDINT := 16#802200;
  DFCid : UINT := 755;
  debounceMethod : USINT := NO_DEBOUNCE;
END_STRUCT;
END_TYPE

TYPE DFC_bds_NoDeb0x8023 : STRUCT
  DTC : UDINT := 16#802300;
  DFCid : UINT := 756;
  debounceMethod : USINT := NO_DEBOUNCE;
END_STRUCT;
END_TYPE

TYPE DFC_bds_NoDeb0x8024 : STRUCT
  DTC : UDINT := 16#802400;
  DFCid : UINT := 757;
  debounceMethod : USINT := NO_DEBOUNCE;
END_STRUCT;
END_TYPE

TYPE DFC_bds_NoDeb0x8025 : STRUCT
  DTC : UDINT := 16#802500;
  DFCid : UINT := 758;
  debounceMethod : USINT := NO_DEBOUNCE;
END_STRUCT;
END_TYPE

TYPE DFC_bds_NoDeb0x8026 : STRUCT
  DTC : UDINT := 16#802600;
  DFCid : UINT := 759;
  debounceMethod : USINT := NO_DEBOUNCE;
END_STRUCT;
END_TYPE

TYPE DFC_bds_NoDeb0x8027 : STRUCT
  DTC : UDINT := 16#802700;
  DFCid : UINT := 760;
  debounceMethod : USINT := NO_DEBOUNCE;
END_STRUCT;
END_TYPE

TYPE DFC_bds_NoDeb0x8028 : STRUCT
  DTC : UDINT := 16#802800;
  DFCid : UINT := 761;
  debounceMethod : USINT := NO_DEBOUNCE;
END_STRUCT;
END_TYPE

TYPE DFC_bds_NoDeb0x8029 : STRUCT
  DTC : UDINT := 16#802900;
  DFCid : UINT := 762;
  debounceMethod : USINT := NO_DEBOUNCE;
END_STRUCT;
END_TYPE

TYPE DFC_bds_NoDeb0x802a : STRUCT
  DTC : UDINT := 16#802A00;
  DFCid : UINT := 763;
  debounceMethod : USINT := NO_DEBOUNCE;
END_STRUCT;
END_TYPE

TYPE DFC_bds_NoDeb0x802b : STRUCT
  DTC : UDINT := 16#802B00;
  DFCid : UINT := 764;
  debounceMethod : USINT := NO_DEBOUNCE;
END_STRUCT;
END_TYPE

TYPE DFC_bds_NoDeb0x802c : STRUCT
  DTC : UDINT := 16#802C00;
  DFCid : UINT := 765;
  debounceMethod : USINT := NO_DEBOUNCE;
END_STRUCT;
END_TYPE

TYPE DFC_bds_NoDeb0x802d : STRUCT
  DTC : UDINT := 16#802D00;
  DFCid : UINT := 766;
  debounceMethod : USINT := NO_DEBOUNCE;
END_STRUCT;
END_TYPE

TYPE DFC_bds_NoDeb0x802e : STRUCT
  DTC : UDINT := 16#802E00;
  DFCid : UINT := 767;
  debounceMethod : USINT := NO_DEBOUNCE;
END_STRUCT;
END_TYPE

TYPE DFC_bds_NoDeb0x802f : STRUCT
  DTC : UDINT := 16#802F00;
  DFCid : UINT := 768;
  debounceMethod : USINT := NO_DEBOUNCE;
END_STRUCT;
END_TYPE

TYPE DFC_bds_NoDeb0x8030 : STRUCT
  DTC : UDINT := 16#803000;
  DFCid : UINT := 769;
  debounceMethod : USINT := NO_DEBOUNCE;
END_STRUCT;
END_TYPE

TYPE DFC_bds_NoDeb0x8031 : STRUCT
  DTC : UDINT := 16#803100;
  DFCid : UINT := 770;
  debounceMethod : USINT := NO_DEBOUNCE;
END_STRUCT;
END_TYPE

TYPE DFC_bds_NoDeb0x8032 : STRUCT
  DTC : UDINT := 16#803200;
  DFCid : UINT := 771;
  debounceMethod : USINT := NO_DEBOUNCE;
END_STRUCT;
END_TYPE

TYPE DFC_bds_NoDeb0x8033 : STRUCT
  DTC : UDINT := 16#803300;
  DFCid : UINT := 772;
  debounceMethod : USINT := NO_DEBOUNCE;
END_STRUCT;
END_TYPE

TYPE DFC_bds_NoDeb0x8034 : STRUCT
  DTC : UDINT := 16#803400;
  DFCid : UINT := 773;
  debounceMethod : USINT := NO_DEBOUNCE;
END_STRUCT;
END_TYPE

TYPE DFC_bds_NoDeb0x8035 : STRUCT
  DTC : UDINT := 16#803500;
  DFCid : UINT := 774;
  debounceMethod : USINT := NO_DEBOUNCE;
END_STRUCT;
END_TYPE

TYPE DFC_bds_NoDeb0x8036 : STRUCT
  DTC : UDINT := 16#803600;
  DFCid : UINT := 775;
  debounceMethod : USINT := NO_DEBOUNCE;
END_STRUCT;
END_TYPE

TYPE DFC_bds_NoDeb0x8037 : STRUCT
  DTC : UDINT := 16#803700;
  DFCid : UINT := 776;
  debounceMethod : USINT := NO_DEBOUNCE;
END_STRUCT;
END_TYPE

TYPE DFC_bds_NoDeb0x8038 : STRUCT
  DTC : UDINT := 16#803800;
  DFCid : UINT := 777;
  debounceMethod : USINT := NO_DEBOUNCE;
END_STRUCT;
END_TYPE

TYPE DFC_bds_NoDeb0x8039 : STRUCT
  DTC : UDINT := 16#803900;
  DFCid : UINT := 778;
  debounceMethod : USINT := NO_DEBOUNCE;
END_STRUCT;
END_TYPE

TYPE DFC_bds_NoDeb0x803a : STRUCT
  DTC : UDINT := 16#803A00;
  DFCid : UINT := 779;
  debounceMethod : USINT := NO_DEBOUNCE;
END_STRUCT;
END_TYPE

TYPE DFC_bds_NoDeb0x803b : STRUCT
  DTC : UDINT := 16#803B00;
  DFCid : UINT := 780;
  debounceMethod : USINT := NO_DEBOUNCE;
END_STRUCT;
END_TYPE

TYPE DFC_bds_NoDeb0x803c : STRUCT
  DTC : UDINT := 16#803C00;
  DFCid : UINT := 781;
  debounceMethod : USINT := NO_DEBOUNCE;
END_STRUCT;
END_TYPE

TYPE DFC_bds_NoDeb0x803d : STRUCT
  DTC : UDINT := 16#803D00;
  DFCid : UINT := 782;
  debounceMethod : USINT := NO_DEBOUNCE;
END_STRUCT;
END_TYPE

TYPE DFC_bds_NoDeb0x803e : STRUCT
  DTC : UDINT := 16#803E00;
  DFCid : UINT := 783;
  debounceMethod : USINT := NO_DEBOUNCE;
END_STRUCT;
END_TYPE

TYPE DFC_bds_NoDeb0x803f : STRUCT
  DTC : UDINT := 16#803F00;
  DFCid : UINT := 784;
  debounceMethod : USINT := NO_DEBOUNCE;
END_STRUCT;
END_TYPE

TYPE DFC_bds_NoDeb0x8040 : STRUCT
  DTC : UDINT := 16#804000;
  DFCid : UINT := 785;
  debounceMethod : USINT := NO_DEBOUNCE;
END_STRUCT;
END_TYPE

TYPE DFC_bds_NoDeb0x8041 : STRUCT
  DTC : UDINT := 16#804100;
  DFCid : UINT := 786;
  debounceMethod : USINT := NO_DEBOUNCE;
END_STRUCT;
END_TYPE

TYPE DFC_bds_NoDeb0x8042 : STRUCT
  DTC : UDINT := 16#804200;
  DFCid : UINT := 787;
  debounceMethod : USINT := NO_DEBOUNCE;
END_STRUCT;
END_TYPE

TYPE DFC_bds_NoDeb0x8043 : STRUCT
  DTC : UDINT := 16#804300;
  DFCid : UINT := 788;
  debounceMethod : USINT := NO_DEBOUNCE;
END_STRUCT;
END_TYPE

TYPE DFC_bds_NoDeb0x8044 : STRUCT
  DTC : UDINT := 16#804400;
  DFCid : UINT := 789;
  debounceMethod : USINT := NO_DEBOUNCE;
END_STRUCT;
END_TYPE

TYPE DFC_bds_NoDeb0x8045 : STRUCT
  DTC : UDINT := 16#804500;
  DFCid : UINT := 790;
  debounceMethod : USINT := NO_DEBOUNCE;
END_STRUCT;
END_TYPE

TYPE DFC_bds_NoDeb0x8046 : STRUCT
  DTC : UDINT := 16#804600;
  DFCid : UINT := 791;
  debounceMethod : USINT := NO_DEBOUNCE;
END_STRUCT;
END_TYPE

TYPE DFC_bds_NoDeb0x8047 : STRUCT
  DTC : UDINT := 16#804700;
  DFCid : UINT := 792;
  debounceMethod : USINT := NO_DEBOUNCE;
END_STRUCT;
END_TYPE

TYPE DFC_bds_NoDeb0x8048 : STRUCT
  DTC : UDINT := 16#804800;
  DFCid : UINT := 793;
  debounceMethod : USINT := NO_DEBOUNCE;
END_STRUCT;
END_TYPE

TYPE DFC_bds_NoDeb0x8049 : STRUCT
  DTC : UDINT := 16#804900;
  DFCid : UINT := 794;
  debounceMethod : USINT := NO_DEBOUNCE;
END_STRUCT;
END_TYPE

TYPE DFC_bds_NoDeb0x804a : STRUCT
  DTC : UDINT := 16#804A00;
  DFCid : UINT := 795;
  debounceMethod : USINT := NO_DEBOUNCE;
END_STRUCT;
END_TYPE

TYPE DFC_bds_NoDeb0x804b : STRUCT
  DTC : UDINT := 16#804B00;
  DFCid : UINT := 796;
  debounceMethod : USINT := NO_DEBOUNCE;
END_STRUCT;
END_TYPE

TYPE DFC_bds_NoDeb0x804c : STRUCT
  DTC : UDINT := 16#804C00;
  DFCid : UINT := 797;
  debounceMethod : USINT := NO_DEBOUNCE;
END_STRUCT;
END_TYPE

TYPE DFC_bds_NoDeb0x804d : STRUCT
  DTC : UDINT := 16#804D00;
  DFCid : UINT := 798;
  debounceMethod : USINT := NO_DEBOUNCE;
END_STRUCT;
END_TYPE

TYPE DFC_bds_NoDeb0x804e : STRUCT
  DTC : UDINT := 16#804E00;
  DFCid : UINT := 799;
  debounceMethod : USINT := NO_DEBOUNCE;
END_STRUCT;
END_TYPE

TYPE DFC_bds_NoDeb0x804f : STRUCT
  DTC : UDINT := 16#804F00;
  DFCid : UINT := 800;
  debounceMethod : USINT := NO_DEBOUNCE;
END_STRUCT;
END_TYPE

TYPE DFC_bds_NoDeb0x8050 : STRUCT
  DTC : UDINT := 16#805000;
  DFCid : UINT := 801;
  debounceMethod : USINT := NO_DEBOUNCE;
END_STRUCT;
END_TYPE

TYPE DFC_bds_NoDeb0x8051 : STRUCT
  DTC : UDINT := 16#805100;
  DFCid : UINT := 802;
  debounceMethod : USINT := NO_DEBOUNCE;
END_STRUCT;
END_TYPE

TYPE DFC_bds_NoDeb0x8052 : STRUCT
  DTC : UDINT := 16#805200;
  DFCid : UINT := 803;
  debounceMethod : USINT := NO_DEBOUNCE;
END_STRUCT;
END_TYPE

TYPE DFC_bds_NoDeb0x8053 : STRUCT
  DTC : UDINT := 16#805300;
  DFCid : UINT := 804;
  debounceMethod : USINT := NO_DEBOUNCE;
END_STRUCT;
END_TYPE

TYPE DFC_bds_NoDeb0x8054 : STRUCT
  DTC : UDINT := 16#805400;
  DFCid : UINT := 805;
  debounceMethod : USINT := NO_DEBOUNCE;
END_STRUCT;
END_TYPE

TYPE DFC_bds_NoDeb0x8055 : STRUCT
  DTC : UDINT := 16#805500;
  DFCid : UINT := 806;
  debounceMethod : USINT := NO_DEBOUNCE;
END_STRUCT;
END_TYPE

TYPE DFC_bds_NoDeb0x8056 : STRUCT
  DTC : UDINT := 16#805600;
  DFCid : UINT := 807;
  debounceMethod : USINT := NO_DEBOUNCE;
END_STRUCT;
END_TYPE

TYPE DFC_bds_NoDeb0x8057 : STRUCT
  DTC : UDINT := 16#805700;
  DFCid : UINT := 808;
  debounceMethod : USINT := NO_DEBOUNCE;
END_STRUCT;
END_TYPE

TYPE DFC_bds_NoDeb0x8058 : STRUCT
  DTC : UDINT := 16#805800;
  DFCid : UINT := 809;
  debounceMethod : USINT := NO_DEBOUNCE;
END_STRUCT;
END_TYPE

TYPE DFC_bds_NoDeb0x8059 : STRUCT
  DTC : UDINT := 16#805900;
  DFCid : UINT := 810;
  debounceMethod : USINT := NO_DEBOUNCE;
END_STRUCT;
END_TYPE

TYPE DFC_bds_NoDeb0x805a : STRUCT
  DTC : UDINT := 16#805A00;
  DFCid : UINT := 811;
  debounceMethod : USINT := NO_DEBOUNCE;
END_STRUCT;
END_TYPE

TYPE DFC_bds_NoDeb0x805b : STRUCT
  DTC : UDINT := 16#805B00;
  DFCid : UINT := 812;
  debounceMethod : USINT := NO_DEBOUNCE;
END_STRUCT;
END_TYPE

TYPE DFC_bds_NoDeb0x805c : STRUCT
  DTC : UDINT := 16#805C00;
  DFCid : UINT := 813;
  debounceMethod : USINT := NO_DEBOUNCE;
END_STRUCT;
END_TYPE

TYPE DFC_bds_NoDeb0x805d : STRUCT
  DTC : UDINT := 16#805D00;
  DFCid : UINT := 814;
  debounceMethod : USINT := NO_DEBOUNCE;
END_STRUCT;
END_TYPE

TYPE DFC_bds_NoDeb0x805e : STRUCT
  DTC : UDINT := 16#805E00;
  DFCid : UINT := 815;
  debounceMethod : USINT := NO_DEBOUNCE;
END_STRUCT;
END_TYPE

TYPE DFC_bds_NoDeb0x805f : STRUCT
  DTC : UDINT := 16#805F00;
  DFCid : UINT := 816;
  debounceMethod : USINT := NO_DEBOUNCE;
END_STRUCT;
END_TYPE

TYPE DFC_bds_NoDeb0x8060 : STRUCT
  DTC : UDINT := 16#806000;
  DFCid : UINT := 817;
  debounceMethod : USINT := NO_DEBOUNCE;
END_STRUCT;
END_TYPE

TYPE DFC_bds_NoDeb0x8061 : STRUCT
  DTC : UDINT := 16#806100;
  DFCid : UINT := 818;
  debounceMethod : USINT := NO_DEBOUNCE;
END_STRUCT;
END_TYPE

TYPE DFC_bds_NoDeb0x8062 : STRUCT
  DTC : UDINT := 16#806200;
  DFCid : UINT := 819;
  debounceMethod : USINT := NO_DEBOUNCE;
END_STRUCT;
END_TYPE

TYPE DFC_bds_NoDeb0x8063 : STRUCT
  DTC : UDINT := 16#806300;
  DFCid : UINT := 106;
  debounceMethod : USINT := TIME_UP_DOWN;
END_STRUCT;
END_TYPE

TYPE DFC_bds_NoDeb0x8064 : STRUCT
  DTC : UDINT := 16#806400;
  DFCid : UINT := 107;
  debounceMethod : USINT := TIME_UP_DOWN;
END_STRUCT;
END_TYPE

TYPE DFC_bds_NoDeb0x8065 : STRUCT
  DTC : UDINT := 16#806500;
  DFCid : UINT := 108;
  debounceMethod : USINT := TIME_UP_DOWN;
END_STRUCT;
END_TYPE

TYPE DFC_bds_NoDeb0x8066 : STRUCT
  DTC : UDINT := 16#806600;
  DFCid : UINT := 109;
  debounceMethod : USINT := TIME_UP_DOWN;
END_STRUCT;
END_TYPE

TYPE DFC_bds_NoDeb0x8067 : STRUCT
  DTC : UDINT := 16#806700;
  DFCid : UINT := 110;
  debounceMethod : USINT := TIME_UP_DOWN;
END_STRUCT;
END_TYPE

TYPE DFC_bds_NoDeb0x8068 : STRUCT
  DTC : UDINT := 16#806800;
  DFCid : UINT := 111;
  debounceMethod : USINT := TIME_UP_DOWN;
END_STRUCT;
END_TYPE

TYPE DFC_bds_NoDeb0x8069 : STRUCT
  DTC : UDINT := 16#806900;
  DFCid : UINT := 112;
  debounceMethod : USINT := TIME_UP_DOWN;
END_STRUCT;
END_TYPE

TYPE DFC_bds_NoDeb0x806a : STRUCT
  DTC : UDINT := 16#806A00;
  DFCid : UINT := 113;
  debounceMethod : USINT := TIME_UP_DOWN;
END_STRUCT;
END_TYPE

TYPE DFC_bds_NoDeb0x806b : STRUCT
  DTC : UDINT := 16#806B00;
  DFCid : UINT := 114;
  debounceMethod : USINT := TIME_UP_DOWN;
END_STRUCT;
END_TYPE

TYPE DFC_bds_NoDeb0x806c : STRUCT
  DTC : UDINT := 16#806C00;
  DFCid : UINT := 115;
  debounceMethod : USINT := TIME_UP_DOWN;
END_STRUCT;
END_TYPE

TYPE DFC_bds_NoDeb0x806d : STRUCT
  DTC : UDINT := 16#806D00;
  DFCid : UINT := 116;
  debounceMethod : USINT := TIME_UP_DOWN;
END_STRUCT;
END_TYPE

TYPE DFC_bds_NoDeb0x806e : STRUCT
  DTC : UDINT := 16#806E00;
  DFCid : UINT := 117;
  debounceMethod : USINT := TIME_UP_DOWN;
END_STRUCT;
END_TYPE

TYPE DFC_bds_NoDeb0x806f : STRUCT
  DTC : UDINT := 16#806F00;
  DFCid : UINT := 118;
  debounceMethod : USINT := TIME_UP_DOWN;
END_STRUCT;
END_TYPE

TYPE DFC_bds_NoDeb0x8070 : STRUCT
  DTC : UDINT := 16#807000;
  DFCid : UINT := 119;
  debounceMethod : USINT := TIME_UP_DOWN;
END_STRUCT;
END_TYPE

TYPE DFC_bds_NoDeb0x8071 : STRUCT
  DTC : UDINT := 16#807100;
  DFCid : UINT := 120;
  debounceMethod : USINT := TIME_UP_DOWN;
END_STRUCT;
END_TYPE

TYPE DFC_bds_NoDeb0x8072 : STRUCT
  DTC : UDINT := 16#807200;
  DFCid : UINT := 121;
  debounceMethod : USINT := TIME_UP_DOWN;
END_STRUCT;
END_TYPE

TYPE DFC_bds_NoDeb0x8073 : STRUCT
  DTC : UDINT := 16#807300;
  DFCid : UINT := 122;
  debounceMethod : USINT := TIME_UP_DOWN;
END_STRUCT;
END_TYPE

TYPE DFC_bds_NoDeb0x8074 : STRUCT
  DTC : UDINT := 16#807400;
  DFCid : UINT := 123;
  debounceMethod : USINT := TIME_UP_DOWN;
END_STRUCT;
END_TYPE

TYPE DFC_bds_NoDeb0x8075 : STRUCT
  DTC : UDINT := 16#807500;
  DFCid : UINT := 124;
  debounceMethod : USINT := TIME_UP_DOWN;
END_STRUCT;
END_TYPE

TYPE DFC_bds_NoDeb0x8076 : STRUCT
  DTC : UDINT := 16#807600;
  DFCid : UINT := 125;
  debounceMethod : USINT := TIME_UP_DOWN;
END_STRUCT;
END_TYPE

TYPE DFC_bds_NoDeb0x8077 : STRUCT
  DTC : UDINT := 16#807700;
  DFCid : UINT := 126;
  debounceMethod : USINT := TIME_UP_DOWN;
END_STRUCT;
END_TYPE

TYPE DFC_bds_NoDeb0x8078 : STRUCT
  DTC : UDINT := 16#807800;
  DFCid : UINT := 127;
  debounceMethod : USINT := TIME_UP_DOWN;
END_STRUCT;
END_TYPE

TYPE DFC_bds_NoDeb0x8079 : STRUCT
  DTC : UDINT := 16#807900;
  DFCid : UINT := 128;
  debounceMethod : USINT := TIME_UP_DOWN;
END_STRUCT;
END_TYPE

TYPE DFC_bds_NoDeb0x807a : STRUCT
  DTC : UDINT := 16#807A00;
  DFCid : UINT := 129;
  debounceMethod : USINT := TIME_UP_DOWN;
END_STRUCT;
END_TYPE

TYPE DFC_bds_NoDeb0x807b : STRUCT
  DTC : UDINT := 16#807B00;
  DFCid : UINT := 130;
  debounceMethod : USINT := TIME_UP_DOWN;
END_STRUCT;
END_TYPE

TYPE DFC_bds_NoDeb0x807c : STRUCT
  DTC : UDINT := 16#807C00;
  DFCid : UINT := 131;
  debounceMethod : USINT := TIME_UP_DOWN;
END_STRUCT;
END_TYPE

TYPE DFC_bds_NoDeb0x807d : STRUCT
  DTC : UDINT := 16#807D00;
  DFCid : UINT := 132;
  debounceMethod : USINT := TIME_UP_DOWN;
END_STRUCT;
END_TYPE

TYPE DFC_bds_NoDeb0x807e : STRUCT
  DTC : UDINT := 16#807E00;
  DFCid : UINT := 133;
  debounceMethod : USINT := TIME_UP_DOWN;
END_STRUCT;
END_TYPE

TYPE DFC_bds_NoDeb0x807f : STRUCT
  DTC : UDINT := 16#807F00;
  DFCid : UINT := 134;
  debounceMethod : USINT := TIME_UP_DOWN;
END_STRUCT;
END_TYPE

TYPE DFC_bds_NoDeb0x8080 : STRUCT
  DTC : UDINT := 16#808000;
  DFCid : UINT := 135;
  debounceMethod : USINT := TIME_UP_DOWN;
END_STRUCT;
END_TYPE

TYPE DFC_bds_NoDeb0x8081 : STRUCT
  DTC : UDINT := 16#808100;
  DFCid : UINT := 136;
  debounceMethod : USINT := TIME_UP_DOWN;
END_STRUCT;
END_TYPE

TYPE DFC_bds_NoDeb0x8082 : STRUCT
  DTC : UDINT := 16#808200;
  DFCid : UINT := 137;
  debounceMethod : USINT := TIME_UP_DOWN;
END_STRUCT;
END_TYPE

TYPE DFC_bds_NoDeb0x8083 : STRUCT
  DTC : UDINT := 16#808300;
  DFCid : UINT := 138;
  debounceMethod : USINT := TIME_UP_DOWN;
END_STRUCT;
END_TYPE

TYPE DFC_bds_NoDeb0x8084 : STRUCT
  DTC : UDINT := 16#808400;
  DFCid : UINT := 139;
  debounceMethod : USINT := TIME_UP_DOWN;
END_STRUCT;
END_TYPE

TYPE DFC_bds_NoDeb0x8085 : STRUCT
  DTC : UDINT := 16#808500;
  DFCid : UINT := 140;
  debounceMethod : USINT := TIME_UP_DOWN;
END_STRUCT;
END_TYPE

TYPE DFC_bds_NoDeb0x8086 : STRUCT
  DTC : UDINT := 16#808600;
  DFCid : UINT := 141;
  debounceMethod : USINT := TIME_UP_DOWN;
END_STRUCT;
END_TYPE

TYPE DFC_bds_NoDeb0x8087 : STRUCT
  DTC : UDINT := 16#808700;
  DFCid : UINT := 142;
  debounceMethod : USINT := TIME_UP_DOWN;
END_STRUCT;
END_TYPE

TYPE DFC_bds_NoDeb0x8088 : STRUCT
  DTC : UDINT := 16#808800;
  DFCid : UINT := 143;
  debounceMethod : USINT := TIME_UP_DOWN;
END_STRUCT;
END_TYPE

TYPE DFC_bds_NoDeb0x8089 : STRUCT
  DTC : UDINT := 16#808900;
  DFCid : UINT := 144;
  debounceMethod : USINT := TIME_UP_DOWN;
END_STRUCT;
END_TYPE

TYPE DFC_bds_NoDeb0x808a : STRUCT
  DTC : UDINT := 16#808A00;
  DFCid : UINT := 145;
  debounceMethod : USINT := TIME_UP_DOWN;
END_STRUCT;
END_TYPE

TYPE DFC_bds_NoDeb0x808b : STRUCT
  DTC : UDINT := 16#808B00;
  DFCid : UINT := 146;
  debounceMethod : USINT := TIME_UP_DOWN;
END_STRUCT;
END_TYPE

TYPE DFC_bds_NoDeb0x808c : STRUCT
  DTC : UDINT := 16#808C00;
  DFCid : UINT := 147;
  debounceMethod : USINT := TIME_UP_DOWN;
END_STRUCT;
END_TYPE

TYPE DFC_bds_NoDeb0x808d : STRUCT
  DTC : UDINT := 16#808D00;
  DFCid : UINT := 148;
  debounceMethod : USINT := TIME_UP_DOWN;
END_STRUCT;
END_TYPE

TYPE DFC_bds_NoDeb0x808e : STRUCT
  DTC : UDINT := 16#808E00;
  DFCid : UINT := 149;
  debounceMethod : USINT := TIME_UP_DOWN;
END_STRUCT;
END_TYPE

TYPE DFC_bds_NoDeb0x808f : STRUCT
  DTC : UDINT := 16#808F00;
  DFCid : UINT := 150;
  debounceMethod : USINT := TIME_UP_DOWN;
END_STRUCT;
END_TYPE

TYPE DFC_bds_NoDeb0x8090 : STRUCT
  DTC : UDINT := 16#809000;
  DFCid : UINT := 151;
  debounceMethod : USINT := TIME_UP_DOWN;
END_STRUCT;
END_TYPE

TYPE DFC_bds_NoDeb0x8091 : STRUCT
  DTC : UDINT := 16#809100;
  DFCid : UINT := 152;
  debounceMethod : USINT := TIME_UP_DOWN;
END_STRUCT;
END_TYPE

TYPE DFC_bds_NoDeb0x8092 : STRUCT
  DTC : UDINT := 16#809200;
  DFCid : UINT := 153;
  debounceMethod : USINT := TIME_UP_DOWN;
END_STRUCT;
END_TYPE

TYPE DFC_bds_NoDeb0x8093 : STRUCT
  DTC : UDINT := 16#809300;
  DFCid : UINT := 154;
  debounceMethod : USINT := TIME_UP_DOWN;
END_STRUCT;
END_TYPE

TYPE DFC_bds_NoDeb0x8094 : STRUCT
  DTC : UDINT := 16#809400;
  DFCid : UINT := 155;
  debounceMethod : USINT := TIME_UP_DOWN;
END_STRUCT;
END_TYPE

TYPE DFC_bds_NoDeb0x8095 : STRUCT
  DTC : UDINT := 16#809500;
  DFCid : UINT := 156;
  debounceMethod : USINT := TIME_UP_DOWN;
END_STRUCT;
END_TYPE

TYPE DFC_bds_NoDeb0x8096 : STRUCT
  DTC : UDINT := 16#809600;
  DFCid : UINT := 157;
  debounceMethod : USINT := TIME_UP_DOWN;
END_STRUCT;
END_TYPE

TYPE DFC_bds_NoDeb0x8097 : STRUCT
  DTC : UDINT := 16#809700;
  DFCid : UINT := 158;
  debounceMethod : USINT := TIME_UP_DOWN;
END_STRUCT;
END_TYPE

TYPE DFC_bds_NoDeb0x8098 : STRUCT
  DTC : UDINT := 16#809800;
  DFCid : UINT := 159;
  debounceMethod : USINT := TIME_UP_DOWN;
END_STRUCT;
END_TYPE

TYPE DFC_bds_NoDeb0x8099 : STRUCT
  DTC : UDINT := 16#809900;
  DFCid : UINT := 160;
  debounceMethod : USINT := TIME_UP_DOWN;
END_STRUCT;
END_TYPE

TYPE DFC_bds_NoDeb0x809a : STRUCT
  DTC : UDINT := 16#809A00;
  DFCid : UINT := 161;
  debounceMethod : USINT := TIME_UP_DOWN;
END_STRUCT;
END_TYPE

TYPE DFC_bds_NoDeb0x809b : STRUCT
  DTC : UDINT := 16#809B00;
  DFCid : UINT := 162;
  debounceMethod : USINT := TIME_UP_DOWN;
END_STRUCT;
END_TYPE

TYPE DFC_bds_NoDeb0x809c : STRUCT
  DTC : UDINT := 16#809C00;
  DFCid : UINT := 163;
  debounceMethod : USINT := TIME_UP_DOWN;
END_STRUCT;
END_TYPE

TYPE DFC_bds_NoDeb0x809d : STRUCT
  DTC : UDINT := 16#809D00;
  DFCid : UINT := 164;
  debounceMethod : USINT := TIME_UP_DOWN;
END_STRUCT;
END_TYPE

TYPE DFC_bds_NoDeb0x809e : STRUCT
  DTC : UDINT := 16#809E00;
  DFCid : UINT := 165;
  debounceMethod : USINT := TIME_UP_DOWN;
END_STRUCT;
END_TYPE

TYPE DFC_bds_NoDeb0x809f : STRUCT
  DTC : UDINT := 16#809F00;
  DFCid : UINT := 166;
  debounceMethod : USINT := TIME_UP_DOWN;
END_STRUCT;
END_TYPE

TYPE DFC_bds_NoDeb0x80a0 : STRUCT
  DTC : UDINT := 16#80A000;
  DFCid : UINT := 167;
  debounceMethod : USINT := TIME_UP_DOWN;
END_STRUCT;
END_TYPE

TYPE DFC_bds_NoDeb0x80a1 : STRUCT
  DTC : UDINT := 16#80A100;
  DFCid : UINT := 168;
  debounceMethod : USINT := TIME_UP_DOWN;
END_STRUCT;
END_TYPE

TYPE DFC_bds_NoDeb0x80a2 : STRUCT
  DTC : UDINT := 16#80A200;
  DFCid : UINT := 169;
  debounceMethod : USINT := TIME_UP_DOWN;
END_STRUCT;
END_TYPE

TYPE DFC_bds_NoDeb0x80a3 : STRUCT
  DTC : UDINT := 16#80A300;
  DFCid : UINT := 170;
  debounceMethod : USINT := TIME_UP_DOWN;
END_STRUCT;
END_TYPE

TYPE DFC_bds_NoDeb0x80a4 : STRUCT
  DTC : UDINT := 16#80A400;
  DFCid : UINT := 171;
  debounceMethod : USINT := TIME_UP_DOWN;
END_STRUCT;
END_TYPE

TYPE DFC_bds_NoDeb0x80a5 : STRUCT
  DTC : UDINT := 16#80A500;
  DFCid : UINT := 172;
  debounceMethod : USINT := TIME_UP_DOWN;
END_STRUCT;
END_TYPE

TYPE DFC_bds_NoDeb0x80a6 : STRUCT
  DTC : UDINT := 16#80A600;
  DFCid : UINT := 173;
  debounceMethod : USINT := TIME_UP_DOWN;
END_STRUCT;
END_TYPE

TYPE DFC_bds_NoDeb0x80a7 : STRUCT
  DTC : UDINT := 16#80A700;
  DFCid : UINT := 174;
  debounceMethod : USINT := TIME_UP_DOWN;
END_STRUCT;
END_TYPE

TYPE DFC_bds_NoDeb0x80a8 : STRUCT
  DTC : UDINT := 16#80A800;
  DFCid : UINT := 175;
  debounceMethod : USINT := TIME_UP_DOWN;
END_STRUCT;
END_TYPE

TYPE DFC_bds_NoDeb0x80a9 : STRUCT
  DTC : UDINT := 16#80A900;
  DFCid : UINT := 176;
  debounceMethod : USINT := TIME_UP_DOWN;
END_STRUCT;
END_TYPE

TYPE DFC_bds_NoDeb0x80aa : STRUCT
  DTC : UDINT := 16#80AA00;
  DFCid : UINT := 177;
  debounceMethod : USINT := TIME_UP_DOWN;
END_STRUCT;
END_TYPE

TYPE DFC_bds_NoDeb0x80ab : STRUCT
  DTC : UDINT := 16#80AB00;
  DFCid : UINT := 178;
  debounceMethod : USINT := TIME_UP_DOWN;
END_STRUCT;
END_TYPE

TYPE DFC_bds_NoDeb0x80ac : STRUCT
  DTC : UDINT := 16#80AC00;
  DFCid : UINT := 179;
  debounceMethod : USINT := TIME_UP_DOWN;
END_STRUCT;
END_TYPE

TYPE DFC_bds_NoDeb0x80ad : STRUCT
  DTC : UDINT := 16#80AD00;
  DFCid : UINT := 180;
  debounceMethod : USINT := TIME_UP_DOWN;
END_STRUCT;
END_TYPE

TYPE DFC_bds_NoDeb0x80ae : STRUCT
  DTC : UDINT := 16#80AE00;
  DFCid : UINT := 181;
  debounceMethod : USINT := TIME_UP_DOWN;
END_STRUCT;
END_TYPE

TYPE DFC_bds_NoDeb0x80af : STRUCT
  DTC : UDINT := 16#80AF00;
  DFCid : UINT := 182;
  debounceMethod : USINT := TIME_UP_DOWN;
END_STRUCT;
END_TYPE

TYPE DFC_bds_NoDeb0x80b0 : STRUCT
  DTC : UDINT := 16#80B000;
  DFCid : UINT := 183;
  debounceMethod : USINT := TIME_UP_DOWN;
END_STRUCT;
END_TYPE

TYPE DFC_bds_NoDeb0x80b1 : STRUCT
  DTC : UDINT := 16#80B100;
  DFCid : UINT := 184;
  debounceMethod : USINT := TIME_UP_DOWN;
END_STRUCT;
END_TYPE

TYPE DFC_bds_NoDeb0x80b2 : STRUCT
  DTC : UDINT := 16#80B200;
  DFCid : UINT := 185;
  debounceMethod : USINT := TIME_UP_DOWN;
END_STRUCT;
END_TYPE

TYPE DFC_bds_NoDeb0x80b3 : STRUCT
  DTC : UDINT := 16#80B300;
  DFCid : UINT := 186;
  debounceMethod : USINT := TIME_UP_DOWN;
END_STRUCT;
END_TYPE

TYPE DFC_bds_NoDeb0x80b4 : STRUCT
  DTC : UDINT := 16#80B400;
  DFCid : UINT := 187;
  debounceMethod : USINT := TIME_UP_DOWN;
END_STRUCT;
END_TYPE

TYPE DFC_bds_NoDeb0x80b5 : STRUCT
  DTC : UDINT := 16#80B500;
  DFCid : UINT := 188;
  debounceMethod : USINT := TIME_UP_DOWN;
END_STRUCT;
END_TYPE

TYPE DFC_bds_NoDeb0x80b6 : STRUCT
  DTC : UDINT := 16#80B600;
  DFCid : UINT := 189;
  debounceMethod : USINT := TIME_UP_DOWN;
END_STRUCT;
END_TYPE

TYPE DFC_bds_NoDeb0x80b7 : STRUCT
  DTC : UDINT := 16#80B700;
  DFCid : UINT := 190;
  debounceMethod : USINT := TIME_UP_DOWN;
END_STRUCT;
END_TYPE

TYPE DFC_bds_NoDeb0x80b8 : STRUCT
  DTC : UDINT := 16#80B800;
  DFCid : UINT := 191;
  debounceMethod : USINT := TIME_UP_DOWN;
END_STRUCT;
END_TYPE

TYPE DFC_bds_NoDeb0x80b9 : STRUCT
  DTC : UDINT := 16#80B900;
  DFCid : UINT := 192;
  debounceMethod : USINT := TIME_UP_DOWN;
END_STRUCT;
END_TYPE

TYPE DFC_bds_NoDeb0x80ba : STRUCT
  DTC : UDINT := 16#80BA00;
  DFCid : UINT := 193;
  debounceMethod : USINT := TIME_UP_DOWN;
END_STRUCT;
END_TYPE

TYPE DFC_bds_NoDeb0x80bb : STRUCT
  DTC : UDINT := 16#80BB00;
  DFCid : UINT := 194;
  debounceMethod : USINT := TIME_UP_DOWN;
END_STRUCT;
END_TYPE

TYPE DFC_bds_NoDeb0x80bc : STRUCT
  DTC : UDINT := 16#80BC00;
  DFCid : UINT := 195;
  debounceMethod : USINT := TIME_UP_DOWN;
END_STRUCT;
END_TYPE

TYPE DFC_bds_NoDeb0x80bd : STRUCT
  DTC : UDINT := 16#80BD00;
  DFCid : UINT := 196;
  debounceMethod : USINT := TIME_UP_DOWN;
END_STRUCT;
END_TYPE

TYPE DFC_bds_NoDeb0x80be : STRUCT
  DTC : UDINT := 16#80BE00;
  DFCid : UINT := 197;
  debounceMethod : USINT := TIME_UP_DOWN;
END_STRUCT;
END_TYPE

TYPE DFC_bds_NoDeb0x80bf : STRUCT
  DTC : UDINT := 16#80BF00;
  DFCid : UINT := 198;
  debounceMethod : USINT := TIME_UP_DOWN;
END_STRUCT;
END_TYPE

TYPE DFC_bds_NoDeb0x80c0 : STRUCT
  DTC : UDINT := 16#80C000;
  DFCid : UINT := 199;
  debounceMethod : USINT := TIME_UP_DOWN;
END_STRUCT;
END_TYPE

TYPE DFC_bds_NoDeb0x80c1 : STRUCT
  DTC : UDINT := 16#80C100;
  DFCid : UINT := 200;
  debounceMethod : USINT := TIME_UP_DOWN;
END_STRUCT;
END_TYPE

TYPE DFC_bds_NoDeb0x80c2 : STRUCT
  DTC : UDINT := 16#80C200;
  DFCid : UINT := 201;
  debounceMethod : USINT := TIME_UP_DOWN;
END_STRUCT;
END_TYPE

TYPE DFC_bds_NoDeb0x80c3 : STRUCT
  DTC : UDINT := 16#80C300;
  DFCid : UINT := 202;
  debounceMethod : USINT := TIME_UP_DOWN;
END_STRUCT;
END_TYPE

TYPE DFC_bds_NoDeb0x80c4 : STRUCT
  DTC : UDINT := 16#80C400;
  DFCid : UINT := 203;
  debounceMethod : USINT := TIME_UP_DOWN;
END_STRUCT;
END_TYPE

TYPE DFC_bds_NoDeb0x80c5 : STRUCT
  DTC : UDINT := 16#80C500;
  DFCid : UINT := 204;
  debounceMethod : USINT := TIME_UP_DOWN;
END_STRUCT;
END_TYPE

TYPE DFC_bds_NoDeb0x80c6 : STRUCT
  DTC : UDINT := 16#80C600;
  DFCid : UINT := 205;
  debounceMethod : USINT := TIME_UP_DOWN;
END_STRUCT;
END_TYPE

TYPE DFC_bds_NoDeb0x80c7 : STRUCT
  DTC : UDINT := 16#80C700;
  DFCid : UINT := 1;
  debounceMethod : USINT := TIME_IN_ROW;
END_STRUCT;
END_TYPE

TYPE DFC_bds_NoDeb0x80c8 : STRUCT
  DTC : UDINT := 16#80C800;
  DFCid : UINT := 2;
  debounceMethod : USINT := TIME_IN_ROW;
END_STRUCT;
END_TYPE

TYPE DFC_bds_NoDeb0x80c9 : STRUCT
  DTC : UDINT := 16#80C900;
  DFCid : UINT := 3;
  debounceMethod : USINT := TIME_IN_ROW;
END_STRUCT;
END_TYPE

TYPE DFC_bds_NoDeb0x80ca : STRUCT
  DTC : UDINT := 16#80CA00;
  DFCid : UINT := 4;
  debounceMethod : USINT := TIME_IN_ROW;
END_STRUCT;
END_TYPE

TYPE DFC_bds_NoDeb0x80cb : STRUCT
  DTC : UDINT := 16#80CB00;
  DFCid : UINT := 5;
  debounceMethod : USINT := TIME_IN_ROW;
END_STRUCT;
END_TYPE

TYPE DFC_bds_NoDeb0x80cc : STRUCT
  DTC : UDINT := 16#80CC00;
  DFCid : UINT := 6;
  debounceMethod : USINT := TIME_IN_ROW;
END_STRUCT;
END_TYPE

TYPE DFC_bds_NoDeb0x80cd : STRUCT
  DTC : UDINT := 16#80CD00;
  DFCid : UINT := 7;
  debounceMethod : USINT := TIME_IN_ROW;
END_STRUCT;
END_TYPE

TYPE DFC_bds_NoDeb0x80ce : STRUCT
  DTC : UDINT := 16#80CE00;
  DFCid : UINT := 8;
  debounceMethod : USINT := TIME_IN_ROW;
END_STRUCT;
END_TYPE

TYPE DFC_bds_NoDeb0x80cf : STRUCT
  DTC : UDINT := 16#80CF00;
  DFCid : UINT := 9;
  debounceMethod : USINT := TIME_IN_ROW;
END_STRUCT;
END_TYPE

TYPE DFC_bds_NoDeb0x80d0 : STRUCT
  DTC : UDINT := 16#80D000;
  DFCid : UINT := 10;
  debounceMethod : USINT := TIME_IN_ROW;
END_STRUCT;
END_TYPE

TYPE DFC_bds_NoDeb0x80d1 : STRUCT
  DTC : UDINT := 16#80D100;
  DFCid : UINT := 11;
  debounceMethod : USINT := TIME_IN_ROW;
END_STRUCT;
END_TYPE

TYPE DFC_bds_NoDeb0x80d2 : STRUCT
  DTC : UDINT := 16#80D200;
  DFCid : UINT := 12;
  debounceMethod : USINT := TIME_IN_ROW;
END_STRUCT;
END_TYPE

TYPE DFC_bds_NoDeb0x80d3 : STRUCT
  DTC : UDINT := 16#80D300;
  DFCid : UINT := 13;
  debounceMethod : USINT := TIME_IN_ROW;
END_STRUCT;
END_TYPE

TYPE DFC_bds_NoDeb0x80d4 : STRUCT
  DTC : UDINT := 16#80D400;
  DFCid : UINT := 14;
  debounceMethod : USINT := TIME_IN_ROW;
END_STRUCT;
END_TYPE

TYPE DFC_bds_NoDeb0x80d5 : STRUCT
  DTC : UDINT := 16#80D500;
  DFCid : UINT := 15;
  debounceMethod : USINT := TIME_IN_ROW;
END_STRUCT;
END_TYPE

TYPE DFC_bds_NoDeb0x80d6 : STRUCT
  DTC : UDINT := 16#80D600;
  DFCid : UINT := 16;
  debounceMethod : USINT := TIME_IN_ROW;
END_STRUCT;
END_TYPE

TYPE DFC_bds_NoDeb0x80d7 : STRUCT
  DTC : UDINT := 16#80D700;
  DFCid : UINT := 17;
  debounceMethod : USINT := TIME_IN_ROW;
END_STRUCT;
END_TYPE

TYPE DFC_bds_NoDeb0x80d8 : STRUCT
  DTC : UDINT := 16#80D800;
  DFCid : UINT := 18;
  debounceMethod : USINT := TIME_IN_ROW;
END_STRUCT;
END_TYPE

TYPE DFC_bds_NoDeb0x80d9 : STRUCT
  DTC : UDINT := 16#80D900;
  DFCid : UINT := 19;
  debounceMethod : USINT := TIME_IN_ROW;
END_STRUCT;
END_TYPE

TYPE DFC_bds_NoDeb0x80da : STRUCT
  DTC : UDINT := 16#80DA00;
  DFCid : UINT := 20;
  debounceMethod : USINT := TIME_IN_ROW;
END_STRUCT;
END_TYPE

TYPE DFC_bds_NoDeb0x80db : STRUCT
  DTC : UDINT := 16#80DB00;
  DFCid : UINT := 21;
  debounceMethod : USINT := TIME_IN_ROW;
END_STRUCT;
END_TYPE

TYPE DFC_bds_NoDeb0x80dc : STRUCT
  DTC : UDINT := 16#80DC00;
  DFCid : UINT := 22;
  debounceMethod : USINT := TIME_IN_ROW;
END_STRUCT;
END_TYPE

TYPE DFC_bds_NoDeb0x80dd : STRUCT
  DTC : UDINT := 16#80DD00;
  DFCid : UINT := 23;
  debounceMethod : USINT := TIME_IN_ROW;
END_STRUCT;
END_TYPE

TYPE DFC_bds_NoDeb0x80de : STRUCT
  DTC : UDINT := 16#80DE00;
  DFCid : UINT := 24;
  debounceMethod : USINT := TIME_IN_ROW;
END_STRUCT;
END_TYPE

TYPE DFC_bds_NoDeb0x80df : STRUCT
  DTC : UDINT := 16#80DF00;
  DFCid : UINT := 25;
  debounceMethod : USINT := TIME_IN_ROW;
END_STRUCT;
END_TYPE

TYPE DFC_bds_NoDeb0x80e0 : STRUCT
  DTC : UDINT := 16#80E000;
  DFCid : UINT := 26;
  debounceMethod : USINT := TIME_IN_ROW;
END_STRUCT;
END_TYPE

TYPE DFC_bds_NoDeb0x80e1 : STRUCT
  DTC : UDINT := 16#80E100;
  DFCid : UINT := 27;
  debounceMethod : USINT := TIME_IN_ROW;
END_STRUCT;
END_TYPE

TYPE DFC_bds_NoDeb0x80e2 : STRUCT
  DTC : UDINT := 16#80E200;
  DFCid : UINT := 28;
  debounceMethod : USINT := TIME_IN_ROW;
END_STRUCT;
END_TYPE

TYPE DFC_bds_NoDeb0x80e3 : STRUCT
  DTC : UDINT := 16#80E300;
  DFCid : UINT := 29;
  debounceMethod : USINT := TIME_IN_ROW;
END_STRUCT;
END_TYPE

TYPE DFC_bds_NoDeb0x80e4 : STRUCT
  DTC : UDINT := 16#80E400;
  DFCid : UINT := 30;
  debounceMethod : USINT := TIME_IN_ROW;
END_STRUCT;
END_TYPE

TYPE DFC_bds_NoDeb0x80e5 : STRUCT
  DTC : UDINT := 16#80E500;
  DFCid : UINT := 31;
  debounceMethod : USINT := TIME_IN_ROW;
END_STRUCT;
END_TYPE

TYPE DFC_bds_NoDeb0x80e6 : STRUCT
  DTC : UDINT := 16#80E600;
  DFCid : UINT := 32;
  debounceMethod : USINT := TIME_IN_ROW;
END_STRUCT;
END_TYPE

TYPE DFC_bds_NoDeb0x80e7 : STRUCT
  DTC : UDINT := 16#80E700;
  DFCid : UINT := 33;
  debounceMethod : USINT := TIME_IN_ROW;
END_STRUCT;
END_TYPE

TYPE DFC_bds_NoDeb0x80e8 : STRUCT
  DTC : UDINT := 16#80E800;
  DFCid : UINT := 34;
  debounceMethod : USINT := TIME_IN_ROW;
END_STRUCT;
END_TYPE

TYPE DFC_bds_NoDeb0x80e9 : STRUCT
  DTC : UDINT := 16#80E900;
  DFCid : UINT := 35;
  debounceMethod : USINT := TIME_IN_ROW;
END_STRUCT;
END_TYPE

TYPE DFC_bds_NoDeb0x80ea : STRUCT
  DTC : UDINT := 16#80EA00;
  DFCid : UINT := 36;
  debounceMethod : USINT := TIME_IN_ROW;
END_STRUCT;
END_TYPE

TYPE DFC_bds_NoDeb0x80eb : STRUCT
  DTC : UDINT := 16#80EB00;
  DFCid : UINT := 37;
  debounceMethod : USINT := TIME_IN_ROW;
END_STRUCT;
END_TYPE

TYPE DFC_bds_NoDeb0x80ec : STRUCT
  DTC : UDINT := 16#80EC00;
  DFCid : UINT := 38;
  debounceMethod : USINT := TIME_IN_ROW;
END_STRUCT;
END_TYPE

TYPE DFC_bds_NoDeb0x80ed : STRUCT
  DTC : UDINT := 16#80ED00;
  DFCid : UINT := 39;
  debounceMethod : USINT := TIME_IN_ROW;
END_STRUCT;
END_TYPE

TYPE DFC_bds_NoDeb0x80ee : STRUCT
  DTC : UDINT := 16#80EE00;
  DFCid : UINT := 40;
  debounceMethod : USINT := TIME_IN_ROW;
END_STRUCT;
END_TYPE

TYPE DFC_bds_NoDeb0x80ef : STRUCT
  DTC : UDINT := 16#80EF00;
  DFCid : UINT := 41;
  debounceMethod : USINT := TIME_IN_ROW;
END_STRUCT;
END_TYPE

TYPE DFC_bds_NoDeb0x80f0 : STRUCT
  DTC : UDINT := 16#80F000;
  DFCid : UINT := 42;
  debounceMethod : USINT := TIME_IN_ROW;
END_STRUCT;
END_TYPE

TYPE DFC_bds_NoDeb0x80f1 : STRUCT
  DTC : UDINT := 16#80F100;
  DFCid : UINT := 43;
  debounceMethod : USINT := TIME_IN_ROW;
END_STRUCT;
END_TYPE

TYPE DFC_bds_NoDeb0x80f2 : STRUCT
  DTC : UDINT := 16#80F200;
  DFCid : UINT := 44;
  debounceMethod : USINT := TIME_IN_ROW;
END_STRUCT;
END_TYPE

TYPE DFC_bds_NoDeb0x80f3 : STRUCT
  DTC : UDINT := 16#80F300;
  DFCid : UINT := 45;
  debounceMethod : USINT := TIME_IN_ROW;
END_STRUCT;
END_TYPE

TYPE DFC_bds_NoDeb0x80f4 : STRUCT
  DTC : UDINT := 16#80F400;
  DFCid : UINT := 46;
  debounceMethod : USINT := TIME_IN_ROW;
END_STRUCT;
END_TYPE

TYPE DFC_bds_NoDeb0x80f5 : STRUCT
  DTC : UDINT := 16#80F500;
  DFCid : UINT := 47;
  debounceMethod : USINT := TIME_IN_ROW;
END_STRUCT;
END_TYPE

TYPE DFC_bds_NoDeb0x80f6 : STRUCT
  DTC : UDINT := 16#80F600;
  DFCid : UINT := 48;
  debounceMethod : USINT := TIME_IN_ROW;
END_STRUCT;
END_TYPE

TYPE DFC_bds_NoDeb0x80f7 : STRUCT
  DTC : UDINT := 16#80F700;
  DFCid : UINT := 49;
  debounceMethod : USINT := TIME_IN_ROW;
END_STRUCT;
END_TYPE

TYPE DFC_bds_NoDeb0x80f8 : STRUCT
  DTC : UDINT := 16#80F800;
  DFCid : UINT := 50;
  debounceMethod : USINT := TIME_IN_ROW;
END_STRUCT;
END_TYPE

TYPE DFC_bds_NoDeb0x80f9 : STRUCT
  DTC : UDINT := 16#80F900;
  DFCid : UINT := 51;
  debounceMethod : USINT := TIME_IN_ROW;
END_STRUCT;
END_TYPE

TYPE DFC_bds_NoDeb0x80fa : STRUCT
  DTC : UDINT := 16#80FA00;
  DFCid : UINT := 52;
  debounceMethod : USINT := TIME_IN_ROW;
END_STRUCT;
END_TYPE

TYPE DFC_bds_NoDeb0x80fb : STRUCT
  DTC : UDINT := 16#80FB00;
  DFCid : UINT := 53;
  debounceMethod : USINT := TIME_IN_ROW;
END_STRUCT;
END_TYPE

TYPE DFC_bds_NoDeb0x80fc : STRUCT
  DTC : UDINT := 16#80FC00;
  DFCid : UINT := 54;
  debounceMethod : USINT := TIME_IN_ROW;
END_STRUCT;
END_TYPE

TYPE DFC_bds_NoDeb0x80fd : STRUCT
  DTC : UDINT := 16#80FD00;
  DFCid : UINT := 55;
  debounceMethod : USINT := TIME_IN_ROW;
END_STRUCT;
END_TYPE

TYPE DFC_bds_NoDeb0x80fe : STRUCT
  DTC : UDINT := 16#80FE00;
  DFCid : UINT := 56;
  debounceMethod : USINT := TIME_IN_ROW;
END_STRUCT;
END_TYPE

TYPE DFC_bds_NoDeb0x80ff : STRUCT
  DTC : UDINT := 16#80FF00;
  DFCid : UINT := 57;
  debounceMethod : USINT := TIME_IN_ROW;
END_STRUCT;
END_TYPE

TYPE DFC_bds_NoDeb0x8100 : STRUCT
  DTC : UDINT := 16#810000;
  DFCid : UINT := 58;
  debounceMethod : USINT := TIME_IN_ROW;
END_STRUCT;
END_TYPE

TYPE DFC_bds_NoDeb0x8101 : STRUCT
  DTC : UDINT := 16#810100;
  DFCid : UINT := 59;
  debounceMethod : USINT := TIME_IN_ROW;
END_STRUCT;
END_TYPE

TYPE DFC_bds_NoDeb0x8102 : STRUCT
  DTC : UDINT := 16#810200;
  DFCid : UINT := 60;
  debounceMethod : USINT := TIME_IN_ROW;
END_STRUCT;
END_TYPE

TYPE DFC_bds_NoDeb0x8103 : STRUCT
  DTC : UDINT := 16#810300;
  DFCid : UINT := 61;
  debounceMethod : USINT := TIME_IN_ROW;
END_STRUCT;
END_TYPE

TYPE DFC_bds_NoDeb0x8104 : STRUCT
  DTC : UDINT := 16#810400;
  DFCid : UINT := 62;
  debounceMethod : USINT := TIME_IN_ROW;
END_STRUCT;
END_TYPE

TYPE DFC_bds_NoDeb0x8105 : STRUCT
  DTC : UDINT := 16#810500;
  DFCid : UINT := 63;
  debounceMethod : USINT := TIME_IN_ROW;
END_STRUCT;
END_TYPE

TYPE DFC_bds_NoDeb0x8106 : STRUCT
  DTC : UDINT := 16#810600;
  DFCid : UINT := 64;
  debounceMethod : USINT := TIME_IN_ROW;
END_STRUCT;
END_TYPE

TYPE DFC_bds_NoDeb0x8107 : STRUCT
  DTC : UDINT := 16#810700;
  DFCid : UINT := 65;
  debounceMethod : USINT := TIME_IN_ROW;
END_STRUCT;
END_TYPE

TYPE DFC_bds_NoDeb0x8108 : STRUCT
  DTC : UDINT := 16#810800;
  DFCid : UINT := 66;
  debounceMethod : USINT := TIME_IN_ROW;
END_STRUCT;
END_TYPE

TYPE DFC_bds_NoDeb0x8109 : STRUCT
  DTC : UDINT := 16#810900;
  DFCid : UINT := 67;
  debounceMethod : USINT := TIME_IN_ROW;
END_STRUCT;
END_TYPE

TYPE DFC_bds_NoDeb0x810a : STRUCT
  DTC : UDINT := 16#810A00;
  DFCid : UINT := 68;
  debounceMethod : USINT := TIME_IN_ROW;
END_STRUCT;
END_TYPE

TYPE DFC_bds_NoDeb0x810b : STRUCT
  DTC : UDINT := 16#810B00;
  DFCid : UINT := 69;
  debounceMethod : USINT := TIME_IN_ROW;
END_STRUCT;
END_TYPE

TYPE DFC_bds_NoDeb0x810c : STRUCT
  DTC : UDINT := 16#810C00;
  DFCid : UINT := 70;
  debounceMethod : USINT := TIME_IN_ROW;
END_STRUCT;
END_TYPE

TYPE DFC_bds_NoDeb0x810d : STRUCT
  DTC : UDINT := 16#810D00;
  DFCid : UINT := 71;
  debounceMethod : USINT := TIME_IN_ROW;
END_STRUCT;
END_TYPE

TYPE DFC_bds_NoDeb0x810e : STRUCT
  DTC : UDINT := 16#810E00;
  DFCid : UINT := 72;
  debounceMethod : USINT := TIME_IN_ROW;
END_STRUCT;
END_TYPE

TYPE DFC_bds_NoDeb0x810f : STRUCT
  DTC : UDINT := 16#810F00;
  DFCid : UINT := 73;
  debounceMethod : USINT := TIME_IN_ROW;
END_STRUCT;
END_TYPE

TYPE DFC_bds_NoDeb0x8110 : STRUCT
  DTC : UDINT := 16#811000;
  DFCid : UINT := 74;
  debounceMethod : USINT := TIME_IN_ROW;
END_STRUCT;
END_TYPE

TYPE DFC_bds_NoDeb0x8111 : STRUCT
  DTC : UDINT := 16#811100;
  DFCid : UINT := 75;
  debounceMethod : USINT := TIME_IN_ROW;
END_STRUCT;
END_TYPE

TYPE DFC_bds_NoDeb0x8112 : STRUCT
  DTC : UDINT := 16#811200;
  DFCid : UINT := 76;
  debounceMethod : USINT := TIME_IN_ROW;
END_STRUCT;
END_TYPE

TYPE DFC_bds_NoDeb0x8113 : STRUCT
  DTC : UDINT := 16#811300;
  DFCid : UINT := 77;
  debounceMethod : USINT := TIME_IN_ROW;
END_STRUCT;
END_TYPE

TYPE DFC_bds_NoDeb0x8114 : STRUCT
  DTC : UDINT := 16#811400;
  DFCid : UINT := 78;
  debounceMethod : USINT := TIME_IN_ROW;
END_STRUCT;
END_TYPE

TYPE DFC_bds_NoDeb0x8115 : STRUCT
  DTC : UDINT := 16#811500;
  DFCid : UINT := 79;
  debounceMethod : USINT := TIME_IN_ROW;
END_STRUCT;
END_TYPE

TYPE DFC_bds_NoDeb0x8116 : STRUCT
  DTC : UDINT := 16#811600;
  DFCid : UINT := 80;
  debounceMethod : USINT := TIME_IN_ROW;
END_STRUCT;
END_TYPE

TYPE DFC_bds_NoDeb0x8117 : STRUCT
  DTC : UDINT := 16#811700;
  DFCid : UINT := 81;
  debounceMethod : USINT := TIME_IN_ROW;
END_STRUCT;
END_TYPE

TYPE DFC_bds_NoDeb0x8118 : STRUCT
  DTC : UDINT := 16#811800;
  DFCid : UINT := 82;
  debounceMethod : USINT := TIME_IN_ROW;
END_STRUCT;
END_TYPE

TYPE DFC_bds_NoDeb0x8119 : STRUCT
  DTC : UDINT := 16#811900;
  DFCid : UINT := 83;
  debounceMethod : USINT := TIME_IN_ROW;
END_STRUCT;
END_TYPE

TYPE DFC_bds_NoDeb0x811a : STRUCT
  DTC : UDINT := 16#811A00;
  DFCid : UINT := 84;
  debounceMethod : USINT := TIME_IN_ROW;
END_STRUCT;
END_TYPE

TYPE DFC_bds_NoDeb0x811b : STRUCT
  DTC : UDINT := 16#811B00;
  DFCid : UINT := 85;
  debounceMethod : USINT := TIME_IN_ROW;
END_STRUCT;
END_TYPE

TYPE DFC_bds_NoDeb0x811c : STRUCT
  DTC : UDINT := 16#811C00;
  DFCid : UINT := 86;
  debounceMethod : USINT := TIME_IN_ROW;
END_STRUCT;
END_TYPE

TYPE DFC_bds_NoDeb0x811d : STRUCT
  DTC : UDINT := 16#811D00;
  DFCid : UINT := 87;
  debounceMethod : USINT := TIME_IN_ROW;
END_STRUCT;
END_TYPE

TYPE DFC_bds_NoDeb0x811e : STRUCT
  DTC : UDINT := 16#811E00;
  DFCid : UINT := 88;
  debounceMethod : USINT := TIME_IN_ROW;
END_STRUCT;
END_TYPE

TYPE DFC_bds_NoDeb0x811f : STRUCT
  DTC : UDINT := 16#811F00;
  DFCid : UINT := 89;
  debounceMethod : USINT := TIME_IN_ROW;
END_STRUCT;
END_TYPE

TYPE DFC_bds_NoDeb0x8120 : STRUCT
  DTC : UDINT := 16#812000;
  DFCid : UINT := 90;
  debounceMethod : USINT := TIME_IN_ROW;
END_STRUCT;
END_TYPE

TYPE DFC_bds_NoDeb0x8121 : STRUCT
  DTC : UDINT := 16#812100;
  DFCid : UINT := 91;
  debounceMethod : USINT := TIME_IN_ROW;
END_STRUCT;
END_TYPE

TYPE DFC_bds_NoDeb0x8122 : STRUCT
  DTC : UDINT := 16#812200;
  DFCid : UINT := 92;
  debounceMethod : USINT := TIME_IN_ROW;
END_STRUCT;
END_TYPE

TYPE DFC_bds_NoDeb0x8123 : STRUCT
  DTC : UDINT := 16#812300;
  DFCid : UINT := 93;
  debounceMethod : USINT := TIME_IN_ROW;
END_STRUCT;
END_TYPE

TYPE DFC_bds_NoDeb0x8124 : STRUCT
  DTC : UDINT := 16#812400;
  DFCid : UINT := 94;
  debounceMethod : USINT := TIME_IN_ROW;
END_STRUCT;
END_TYPE

TYPE DFC_bds_NoDeb0x8125 : STRUCT
  DTC : UDINT := 16#812500;
  DFCid : UINT := 95;
  debounceMethod : USINT := TIME_IN_ROW;
END_STRUCT;
END_TYPE

TYPE DFC_bds_NoDeb0x8126 : STRUCT
  DTC : UDINT := 16#812600;
  DFCid : UINT := 96;
  debounceMethod : USINT := TIME_IN_ROW;
END_STRUCT;
END_TYPE

TYPE DFC_bds_NoDeb0x8127 : STRUCT
  DTC : UDINT := 16#812700;
  DFCid : UINT := 97;
  debounceMethod : USINT := TIME_IN_ROW;
END_STRUCT;
END_TYPE

TYPE DFC_bds_NoDeb0x8128 : STRUCT
  DTC : UDINT := 16#812800;
  DFCid : UINT := 98;
  debounceMethod : USINT := TIME_IN_ROW;
END_STRUCT;
END_TYPE

TYPE DFC_bds_NoDeb0x8129 : STRUCT
  DTC : UDINT := 16#812900;
  DFCid : UINT := 99;
  debounceMethod : USINT := TIME_IN_ROW;
END_STRUCT;
END_TYPE

TYPE DFC_bds_NoDeb0x812a : STRUCT
  DTC : UDINT := 16#812A00;
  DFCid : UINT := 100;
  debounceMethod : USINT := TIME_IN_ROW;
END_STRUCT;
END_TYPE

VAR_GLOBAL  (* GVL_debounceMethod *)
  TIME_IN_ROW : USINT := 0;
  EVENT_IN_ROW : USINT := 1;
  TIME_UP_DOWN : USINT := 2;
  EVENT_UP_DOWN : USINT := 3;
  TIME_UP_DOWN_SMALL : USINT := 4;
  EVENT_UP_DOWN_SMALL : USINT := 5;
  TIME_IN_ROW_SMALL : USINT := 6;
  EVENT_IN_ROW_SMALL : USINT := 7;
  NO_DEBOUNCE : USINT := 8;
  NATIVE : USINT := 8;
END_VAR
